(* IEC 61131-3 sources: daoli-st-library/DL_Algo (part 24) *)

(* ---- FB_DL_FoulingResistanceEstimator.st ---- *)
(*==============================================================================
 * 组件名称 (Component)  : FB_DL_FoulingResistanceEstimator
 * 所属子库 (Sublibrary) : DL_Algo
 * 当前版本 (Version)    : 1.0.0
 * 组件分类 (Category)   : 功能块（FUNCTION_BLOCK）· 换热器本体退化算法底座
 * 兼容性   (Platform)   : CODESYS 3.5 / TwinCAT 3 / 汇川 InoProShop / Schneider Machine Expert
 *                         仅依赖 Standard.library（R_TRIG / LN / ABS / MIN / MAX / LIMIT），零厂商方言
 * 接口依赖 (Depends)    : E_DL_Ne107Status —— 唯一属主为 DL_Device 子库的契约件
 *                         I_DL_DeviceHealth（R13 泳道 A1）。本文件只按成员名引用该枚举，
 *                         不重复定义枚举体（重复定义即同名异型，R33 家族超集风险）。
 * 功能描述 (Function)   : 由热侧/冷侧进出口温度与体积流量算出换热量 Q、对数平均温差
 *                         LMTD 与实测传热系数 K，再由 K 与清洁态基准 K_clean 反算污垢
 *                         热阻 Rf = 1/K − 1/K_clean；在趋势窗 tWindow 内用最小二乘做
 *                         Rf 对时间的线性拟合，输出增长斜率与清洗建议。
 *                         本件是「换热器污垢趋势」工艺件的算法底座：只做「算一个值 +
 *                         算一个趋势」，不判工艺合格、不控阀门、不做结垢成分分析。
 * 边界     (Boundary)   : ① 不做 PID、不做阀门/泵控制；② 不做结垢成分与化学分析；
 *                         ③ 数据不可信（温差过小 / 流量过低 / 两侧热负荷不平衡 /
 *                            输入非有限）时**拒绝更新**并保持上次有效值 —— 宁可不给
 *                            数，也不给脏数（R42 精神：判可用与取值同拍）；
 *                         ④ 不内置换热器几何模型与介质物性库，fCp/fRho 与 K_clean 全部
 *                            由调用方按设备台账注入。
 * 分层声明 (Layer)      : 算法层（DL_Algo）。上游为工艺台账件与 HMI 趋势，下游仅
 *                         Standard.library。零全局变量表引用、零外部变量声明、零物理 IO。
 * 段序     (Segments)   : 段1 实例无条件刷新 → 段2 复位通道（CASE 之前，R39）→
 *                         段3 参数闸门与输入防御 → 段4 数据质量四判据 → 段5 状态机 →
 *                         段6 有效更新与趋势累计 → 段7 结论仲裁 → 段8 码位单一优先级链 →
 *                         段9 出口钳位与保持语义重写。
 * 枚举映射表 (R31)      : eIdle(0)→标签 0｜eValid(10)→标签 10｜eTrend(20)→标签 20｜
 *                         eAdvice(30)→标签 30｜eFault(99)→标签 99。每个成员有且仅有一个
 *                         显式标签，ELSE 只接脏值（2212）。
 * 单拍标志清单 (R25)    : 本件唯一的沿输入是 bReset（复位），其消费点为段2 复位通道。
 *                         预清零点：段1 末（_bResetEdge := _fbTrigReset.Q 每次覆盖）；
 *                         置位点：段1 的 _fbTrigReset 实例调用；自清点：紧随实例调用之后
 *                         的 _bResetEdge 赋值行（下拍 R_TRIG.Q 转假即自然清）。
 * 保持位清单 (R27)      : bCleanAdvice（清洗建议，逐拍由 _bCleanLatched 重写）｜
 *                         fQ / fLmtd / fK / fRf（上次有效值，逐拍由 _fXxxHeld 重写并钳位）｜
 *                         fRfSlope（上次窗口斜率，逐拍重写）。复位沿清除锁存与保持值。
 * 定时器清单 (R40)      : 无 TON/TOF 实例。趋势窗以引脚 tSamplePeriod 累加计时，
 *                         窗边界显式重装基准（_fWinElapsedH := 0），不存在跨窗恒真输入；
 *                         时长到**或**样本数触顶（64）即结算并重开新窗，触顶提前结算是为了
 *                         避免「为了凑时长而丢掉分辨率」，也避免样本触顶后窗永远关不上。
 * 三元一致表 (R35)      : 流量比例守卫 0.05~0.9 / 封顶 0.9 / 判据 `<`（低于即不更新）｜
 *                         热平衡容差守卫 0.02~0.5 / 封顶 0.5 / 判据 `>`（超出即不更新）｜
 *                         最小温差守卫 0.5~20 K / 封顶 20 K / 判据 `<`（低于即不更新）。
 * 镜像量清单 (R38)      : 实时量 fFlowHot / fFlowCold 的唯一消费点是段4 的流量比例
 *                         判定（自学习参考流量 _fFlowHotMax / _fFlowColdMax 在同段更新）；
 *                         本件不设「锁存副本 + 实时镜像」双源，边界量全部取自本拍单次读取。
 * 开源溯源 (Origin)     : 原创实现（参考 OSCAT Building 的「温度/流量进 → 传热系数与
 *                         污垢热阻出」行为定义组织方式，T1-2；OSCAT 现行版为 EPL-2.0，
 *                         归档旧件仍受其原始许可约束 —— 本件只取行为定义与引脚组织，
 *                         未下载库文件、未复制任何源码行，公式取自公开传热学常识：
 *                         Q = m·cp·ΔT、逆/顺流 LMTD、Rf = 1/K − 1/K_clean）。
 *                         许可证结论：无代码复制，本文件为本库原创，随本库许可证发布。
 * 验收向量 (Acceptance) :
 *   V1 热侧 90/70 ℃、冷侧 20/40 ℃、逆流、两侧 10 m³/h：ΔT1 = 90−40 = 50 K、
 *      ΔT2 = 70−20 = 50 K，两温差相等时 LMTD 退化为算术平均 50.0 K；fQ ≈ 232.2 kW
 *      （10 m³/h × 1000 kg/m³ × 4.18 kJ/(kg·K) × 20 K / 3600）。规格记 49.7 K 与
 *      232 kW 为取整口径，本件按上式复算（见偏离留档②）。
 *   V2 fK = 1000、fKClean = 2000 → fRf = 1/1000 − 1/2000 = 5.0E-4 ≥ 3.0E-4 →
 *      bCleanAdvice = TRUE（保持态逐拍重写）。
 *   V3（V-A 除零）fArea = 0 → 16#0002_2210，fK 保持上次值并夹进 ≥ 0（R43）。
 *   V4（V-C 跨拍复验）进入 eTrend 后当拍流量骤降 → 段4 本拍复验流量门限失败 →
 *      本拍不更新、不累计斜率样本（绝不用上一相结论直接算斜率，R42）。
 *   V5（V-D 首拍）上电首拍 bValid = FALSE、fRf = 0.0，且首拍样本**不**写入趋势基准
 *      （R19：首扫只装基准，不参与斜率）。
 * 偏离留档 (Deviation)  :
 *   ① 「流量低于额定比例」的额定量：规格未给出额定流量引脚。本件以块内自学习的
 *      「投运以来观测到的最大流量」为参考（_fFlowHotMax / _fFlowColdMax），比例 =
 *      本拍流量 / 参考流量。理由：不新增引脚即可表达「相对自身额定」的语义；影响：
 *      上电初期参考流量偏低，门限自然宽松，随运行收敛（首拍样本不受门限影响）。
 *   ② V1 的 LMTD 数值：等温差时 LMTD 退化为算术平均（数值稳定性要求），与规格
 *      49.7 K 的取整口径相差 0.3 K，属口径差异而非算法差异，此处显式留档。
 *   ③ 输入非有限与「面积/清洁 K 非正」共用 16#0002_2210（规格故障表只给 3 个故障码，
 *      不新增码位；码位表以 §3.0 为准，编码者不得自行偏移）。
 * 修订历史 (Revision)   :
 *   2026-11-15  v1.0.0  首版入库（Round 13 · 泳道 C · DL_Algo 第 28 件）
 *============================================================================*)

(*-----------------------------------------------------------------------------
 * 枚举: E_DL_FoulingState（归属 FB_DL_FoulingResistanceEstimator，同文件发布）
 *----------------------------------------------------------------------------*)
TYPE E_DL_FoulingState :
(
    eIdle   := 0,    // 空闲：未使能或参数未就绪 / Idle, disabled or parameters not ready
    eValid  := 10,   // 有效：本拍已算出可信的 K 与 Rf / Valid, trustworthy K and Rf computed
    eTrend  := 20,   // 趋势：窗内样本数已达 3，斜率可算 / Trend, at least three window samples
    eAdvice := 30,   // 建议清洗：热阻或其斜率越阈（锁存）/ Cleaning advised, latched
    eFault  := 99    // 故障：参数非法或输入非有限 / Fault, illegal parameter or non-finite input
) UINT;
END_TYPE

FUNCTION_BLOCK FB_DL_FoulingResistanceEstimator
VAR_INPUT
    bEnable         : BOOL;                 // 使能（Enable），FALSE = 冻结更新并回空闲；复位通道不受其屏蔽 / Enable, FALSE freezes updates
    bReset          : BOOL;                 // 复位（Reset），上升沿清趋势窗、清洗锁存与保持值 / Rising edge clears trend window and latches
    fTinHot         : REAL;                 // 热侧进口温度（Hot inlet temperature）[℃]，域 −50~300 / Hot side inlet temperature [degC]
    fToutHot        : REAL;                 // 热侧出口温度（Hot outlet temperature）[℃]，域 −50~300 / Hot side outlet temperature [degC]
    fTinCold        : REAL;                 // 冷侧进口温度（Cold inlet temperature）[℃]，域 −50~300 / Cold side inlet temperature [degC]
    fToutCold       : REAL;                 // 冷侧出口温度（Cold outlet temperature）[℃]，域 −50~300 / Cold side outlet temperature [degC]
    fFlowHot        : REAL;                 // 热侧体积流量（Hot volumetric flow）[m³/h]，域 0~10000 / Hot volumetric flow [m3/h]
    fFlowCold       : REAL;                 // 冷侧体积流量（Cold volumetric flow）[m³/h]，域 0~10000 / Cold volumetric flow [m3/h]
    fCpHot          : REAL := 4.18;         // 热侧比热（Hot specific heat）[kJ/(kg·K)]，域 0.5~10，默认 4.18 / Hot specific heat [kJ/(kg K)]
    fCpCold         : REAL := 4.18;         // 冷侧比热（Cold specific heat）[kJ/(kg·K)]，域 0.5~10，默认 4.18 / Cold specific heat [kJ/(kg K)]
    fRhoHot         : REAL := 1000.0;       // 热侧密度（Hot density）[kg/m³]，域 1~2000，默认 1000.0 / Hot density [kg/m3]
    fRhoCold        : REAL := 1000.0;       // 冷侧密度（Cold density）[kg/m³]，域 1~2000，默认 1000.0 / Cold density [kg/m3]
    fArea           : REAL;                 // 换热面积（Heat transfer area）[m²]，域 >0，除零保护对象 / Heat transfer area [m2], must be positive
    fKClean         : REAL;                 // 清洁态传热系数基准（Clean-condition K）[W/(m²·K)]，域 >0 / Clean-condition K [W/(m2 K)], must be positive
    bCounterFlow    : BOOL := TRUE;         // 流型（Flow arrangement），TRUE = 逆流，FALSE = 顺流，默认 TRUE / TRUE counter-flow, FALSE parallel-flow
    fDtmMin         : REAL := 2.0;          // 最小可用温差（Minimum usable temperature difference）[K]，域 0.5~20，默认 2.0 / Minimum usable LMTD [K]
    fHeatBalTol     : REAL := 0.10;         // 两侧热负荷允许偏差比（Heat balance tolerance）[-]，域 0.02~0.5，默认 0.10 / Heat balance tolerance [-]
    fFlowMinRatio   : REAL := 0.20;         // 流量下限比例（Minimum flow ratio）[-]，域 0.05~0.9，默认 0.20 / Minimum flow ratio [-]
    tWindow         : TIME := T#1H;         // 趋势窗长（Trend window），域 5 min~24 h，默认 1 h / Trend window, default 1 h
    tSamplePeriod   : TIME := T#10S;        // 调用周期（Call period）[ms]，必须与实际任务周期一致，默认 10 s / Call period, must match the task
    fRfAlarm        : REAL := 3.0E-4;       // 污垢热阻报警阈（Fouling resistance alarm）[m²·K/W]，域 1E-5~5E-3 / Fouling resistance alarm [m2 K/W]
    fSlopeAlarm     : REAL := 2.0E-5;       // 污垢增长速率阈（Fouling slope alarm）[m²·K/(W·h)]，域 1E-7~1E-3 / Fouling slope alarm [m2 K/(W h)]
END_VAR

VAR_OUTPUT
    fQ              : REAL;                 // 热负荷两侧平均（Heat duty, mean of both sides）[kW]，保持语义 / Mean heat duty of both sides [kW], held
    fLmtd           : REAL;                 // 对数平均温差（Log mean temperature difference）[K]，保持语义 / LMTD [K], held
    fK              : REAL;                 // 实测传热系数（Measured overall K）[W/(m²·K)]，保持语义且夹进 ≥0 / Measured K [W/(m2 K)], held and clamped non-negative
    fRf             : REAL;                 // 污垢热阻（Fouling resistance）[m²·K/W]，= 1/K − 1/K_clean，保持语义 / Fouling resistance [m2 K/W], held
    fRfSlope        : REAL;                 // 窗内趋势斜率（Trend slope in window）[m²·K/(W·h)]，保持语义 / Trend slope [m2 K/(W h)], held
    bValid          : BOOL;                 // 本拍输出有效（Output valid this scan），数据质量不足时为 FALSE / TRUE when this scan produced a trustworthy value
    bCleanAdvice    : BOOL;                 // 建议清洗（Cleaning advised），保持语义（R27），复位沿清除 / Cleaning advised, held until reset
    eHealth         : E_DL_Ne107Status;     // 健康态（NE107 health），引用属主 A1 的枚举 / NE107 health state, owned by A1
    uDiagCode       : UDINT;                // 诊断码（Diagnostic code），本拍单一优先级链输出 / Diagnostic code, single priority chain
    uErrorId        : UDINT;                // 故障码（Error code），仅故障级码，0 = 无故障 / Fault-level code, 0 = no fault
    bError          : BOOL;                 // 故障标志（Error），仅故障级码置位，信息级不置位 / TRUE only for fault-level codes
    nUpdateCount    : UDINT;                // 有效更新次数（Valid update counter）[次]，每次有效更新 +1 / Valid update counter [count]
END_VAR

VAR
    _eState         : E_DL_FoulingState := E_DL_FoulingState.eIdle; // 内部状态（Internal state）/ Internal state machine value
    _bInit          : BOOL;                 // 首扫标志（First-scan flag），初值 FALSE，唯一首扫判据为 NOT _bInit（R19）/ First-scan flag, FALSE by default
    _bSkipSample    : BOOL;                 // 本拍不参与斜率（Skip trend sample this scan），首扫与不可信拍置位 / Skip this scan as a trend sample
    _bParamOk       : BOOL;                 // 参数闸门通过（Parameter gate passed）/ Parameter gate result
    _bDataOk        : BOOL;                 // 数据质量通过（Data quality passed）/ Data quality result
    _bValidNow      : BOOL;                 // 本拍有效（Valid this scan）/ Valid this scan
    _bFaultCond     : BOOL;                 // 故障条件（Fault condition latch-free flag）/ Fault condition flag
    _uFaultCode     : UDINT;                // 本拍故障级码（Fault-level code this scan）/ Fault-level code of this scan
    _uFaultLatched  : UDINT;                // 故障码锁存（Latched fault code），仅复位沿清除 / Latched fault code, reset only
    _uInfoCode      : UDINT;                // 本拍信息级码（Info-level code this scan），每拍重算 / Info-level code, recomputed every scan
    _bArrPrev       : BOOL;                 // 上拍流型（Previous flow arrangement）/ Flow arrangement of the previous scan
    _bArrKnown      : BOOL;                 // 流型已记录（Arrangement recorded）/ Arrangement recorded flag
    _fAreaEff       : REAL;                 // 生效换热面积（Effective area）[m²]，闸门后值 / Effective area [m2] after the gate
    _fKCleanEff     : REAL;                 // 生效清洁 K（Effective clean K）[W/(m²·K)] / Effective clean K [W/(m2 K)]
    _fDtmMinEff     : REAL;                 // 生效最小温差（Effective minimum LMTD）[K]，钳位 0.5~20 / Effective minimum LMTD [K], clamped
    _fBalTolEff     : REAL;                 // 生效热平衡容差（Effective heat balance tolerance）[-]，钳位 0.02~0.5 / Effective heat balance tolerance, clamped
    _fFlowRatioEff  : REAL;                 // 生效流量比例（Effective minimum flow ratio）[-]，钳位 0.05~0.9 / Effective minimum flow ratio, clamped
    _fFlowHotMax    : REAL;                 // 热侧参考流量（Hot reference flow）[m³/h]，自学习峰值 / Self-learned hot reference flow [m3/h]
    _fFlowColdMax   : REAL;                 // 冷侧参考流量（Cold reference flow）[m³/h]，自学习峰值 / Self-learned cold reference flow [m3/h]
    _fQHot          : REAL;                 // 热侧放热量（Heat duty, hot side）[kW]，有符号 / Hot-side duty [kW], signed
    _fQCold         : REAL;                 // 冷侧吸热量（Heat duty, cold side）[kW]，有符号 / Cold-side duty [kW], signed
    _fQMean         : REAL;                 // 两侧平均热负荷（Mean duty）[kW] / Mean duty of both sides [kW]
    _fDt1           : REAL;                 // 端差一（Terminal difference one）[K]，按流型取 / Terminal temperature difference one [K]
    _fDt2           : REAL;                 // 端差二（Terminal difference two）[K]，按流型取 / Terminal temperature difference two [K]
    _fLmtdCalc      : REAL;                 // 本拍 LMTD 计算值（Computed LMTD）[K] / Computed LMTD [K]
    _fLmtdAbs       : REAL;                 // 端差差值的绝对值（Absolute terminal difference gap）[K]，退化判据 / Absolute gap between terminal differences [K]
    _fLmtdDen       : REAL;                 // 对数比值（Logarithmic ratio）[-]，除零保护对象 / Logarithmic ratio, divide-guard object
    _fBalDev        : REAL;                 // 热平衡偏差比（Heat balance deviation）[-] / Heat balance deviation ratio [-]
    _fBalRef        : REAL;                 // 热平衡参考量（Heat balance reference）[kW]/ Reference magnitude for the balance test [kW]
    _fKCalc         : REAL;                 // 本拍 K 计算值（Computed K）[W/(m²·K)] / Computed K [W/(m2 K)]
    _fRfCalc        : REAL;                 // 本拍 Rf 计算值（Computed Rf）[m²·K/W] / Computed Rf [m2 K/W]
    _fQHeld         : REAL;                 // 保持的热负荷（Held heat duty）[kW] / Held heat duty [kW]
    _fLmtdHeld      : REAL;                 // 保持的 LMTD（Held LMTD）[K] / Held LMTD [K]
    _fKHeld         : REAL;                 // 保持的 K（Held K）[W/(m²·K)] / Held K [W/(m2 K)]
    _fRfHeld        : REAL;                 // 保持的 Rf（Held Rf）[m²·K/W] / Held Rf [m2 K/W]
    _fSlopeHeld     : REAL;                 // 保持的斜率（Held slope）[m²·K/(W·h)] / Held slope [m2 K/(W h)]
    _bCleanLatched  : BOOL;                 // 清洗建议锁存（Cleaning advice latch），仅复位沿清除 / Cleaning advice latch, reset only
    _nWinN          : INT;                  // 窗内样本数（Window sample count）[个]，上限 64 / Window sample count, capped at 64
    _fWinElapsedH   : REAL;                 // 窗内已历时（Elapsed hours in window）[h] / Elapsed hours in the current window [h]
    _fWinX          : REAL;                 // 最小二乘 Σt（Sum of time stamps）[h] / Least-squares sum of time stamps [h]
    _fWinY          : REAL;                 // 最小二乘 ΣRf（Sum of Rf samples）[m²·K/W] / Least-squares sum of Rf samples [m2 K/W]
    _fWinXY         : REAL;                 // 最小二乘 Σt·Rf（Sum of products）[h·m²·K/W] / Least-squares sum of products
    _fWinXX         : REAL;                 // 最小二乘 Σt²（Sum of squared times）[h²] / Least-squares sum of squared times [h2]
    _fWinDen        : REAL;                 // 最小二乘分母（Normal-equation denominator）[-]，除零保护对象 / Denominator of the normal equations
    _fWinNum        : REAL;                 // 最小二乘分子（Normal-equation numerator）[-] / Numerator of the normal equations
    _fDtHours       : REAL;                 // 本拍步长（Step in hours）[h]，由 tSamplePeriod 折算 / Step in hours, derived from the call period
    _fWinHoursEff   : REAL;                 // 生效窗长（Effective window length）[h]，由 tWindow 折算 / Effective window length [h]
    _fbTrigReset    : R_TRIG;               // 复位沿（Reset edge detector），主体最前部无条件刷新 / Reset edge detector, refreshed unconditionally
    _bResetEdge     : BOOL;                 // 复位沿单拍标志（Reset one-shot flag），紧随实例自清 / Reset one-shot flag, cleared right after the call
END_VAR

VAR CONSTANT
    DL_FRE_REAL_MAX   : REAL := 3.4E38;      // 单精度有限值判据幅值（Finite magnitude bound）/ Finite bound for REAL inputs
    DL_FRE_EPS        : REAL := 1.0E-6;      // 浮点防零容差（Divide-guard epsilon）/ Float divide-guard epsilon
    DL_FRE_K_MAX      : REAL := 1.0E9;       // K 出口上限（K output ceiling）[W/(m²·K)] / Upper clamp of K [W/(m2 K)]
    DL_FRE_RF_MAX     : REAL := 1.0;         // Rf 出口上限（Rf output ceiling）[m²·K/W] / Upper clamp of Rf [m2 K/W]
    DL_FRE_SLOPE_MAX  : REAL := 1.0;         // 斜率出口上限（Slope output ceiling）[m²·K/(W·h)] / Upper clamp of slope
    DL_FRE_SLOPE_MIN  : REAL := -1.0;        // 斜率出口下限（Slope output floor）[m²·K/(W·h)] / Lower clamp of slope
    DL_FRE_WIN_MAX    : INT  := 64;          // 窗内样本上限（Window sample ceiling）[个] / Window sample ceiling
    DL_FRE_MS_PER_H   : REAL := 3600000.0;   // 毫秒→小时换算（Milliseconds-to-hours scale）[-] / Milliseconds-to-hours scale
    DL_FRE_KW_SCALE   : REAL := 3600.0;      // m³/h·kg/m³·kJ/(kg·K)·K → kW 的换算（Duty unit scale）[-] / Duty unit scale
    DL_FRE_W_SCALE    : REAL := 1000.0;      // kW → W 换算（Kilowatt-to-watt scale）[-] / Kilowatt-to-watt scale
    DL_FRE_DTM_MIN    : REAL := 0.5;         // 最小温差域下限（Minimum LMTD lower clamp）[K] / Minimum LMTD lower clamp [K]
    DL_FRE_DTM_MAX    : REAL := 20.0;        // 最小温差域上限（Minimum LMTD upper clamp）[K] / Minimum LMTD upper clamp [K]
    DL_FRE_TOL_MIN    : REAL := 0.02;        // 热平衡容差域下限（Balance tolerance lower clamp）[-] / Balance tolerance lower clamp
    DL_FRE_TOL_MAX    : REAL := 0.5;         // 热平衡容差域上限（Balance tolerance upper clamp）[-] / Balance tolerance upper clamp
    DL_FRE_RATIO_MIN  : REAL := 0.05;        // 流量比例域下限（Flow ratio lower clamp）[-] / Flow ratio lower clamp
    DL_FRE_RATIO_MAX  : REAL := 0.9;         // 流量比例域上限（Flow ratio upper clamp）[-] / Flow ratio upper clamp
    DL_FRE_RF_FLOOR   : REAL := 0.0;         // Rf 出口下限（Rf output floor）[m²·K/W]，K>K_clean 时按 0 / Rf floor, zero when K exceeds clean K
    DL_FRE_WIN_MIN_N  : INT  := 3;           // 斜率所需最少样本（Minimum samples for a slope）[个] / Minimum samples for the slope
    DL_FRE_ERR_PARAM  : UDINT := 16#0002_2210; // 0002_2210 面积/清洁 K 非正或输入非有限【故障级】/ Illegal area, clean K or non-finite input
    DL_FRE_ERR_LMTD   : UDINT := 16#0002_2211; // 0002_2211 LMTD ≤ 0（温度交叉或流型用错）【故障级】/ Non-positive LMTD
    DL_FRE_ERR_STATE  : UDINT := 16#0002_2212; // 0002_2212 非法状态兜底【故障级】/ Illegal state fallback
    DL_FRE_INFO_LMTD  : UDINT := 16#0002_2201; // 0002_2201 LMTD 低于最小可用温差【信息级】/ LMTD below the usable limit
    DL_FRE_INFO_FLOW  : UDINT := 16#0002_2202; // 0002_2202 流量低于下限比例【信息级】/ Flow below the minimum ratio
    DL_FRE_INFO_BAL   : UDINT := 16#0002_2203; // 0002_2203 两侧热负荷偏差超容差【信息级】/ Heat balance exceeded
    DL_FRE_INFO_ARR   : UDINT := 16#0002_2204; // 0002_2204 逆/顺流口径切换，趋势基准已重置【信息级】/ Arrangement changed, trend reset
END_VAR

// ============================================================================
// 段 1｜实例无条件周期刷新（R7/0.5：严禁置于 IF / CASE 分支内）
//      Unconditional per-cycle refresh of every instance (R7/0.5)
// ============================================================================
_fbTrigReset(CLK := bReset);            // 复位沿实例调用（Reset edge instance call）
_bResetEdge := _fbTrigReset.Q;          // 单拍标志紧随实例赋值，下拍自然清（R24/R25 自清点）

// 本拍故障/信息码与结论预置（每拍重算，杜绝跨拍残留）
// Per-scan preset of codes and conclusions, no cross-scan residue
_uFaultCode  := _uFaultLatched;         // 故障码以上拍锁存续用（Carry the latched fault code）
_uInfoCode   := 16#0000_0000;           // 信息级码预清零（Info code preset to zero）
_bFaultCond  := FALSE;                  // 故障条件预清零（Fault condition preset FALSE）
_bParamOk    := FALSE;                  // 参数闸门预置未通过（Parameter gate preset closed）
_bDataOk     := FALSE;                  // 数据质量预置未通过（Data quality preset failed）
_bValidNow   := FALSE;                  // 本拍有效预置假（Valid preset FALSE）
_bSkipSample := FALSE;                  // 采样跳过预置假（Sample skip preset FALSE）

// 调用周期折算为小时，非法周期按复位通道外的钳位处理（不做除零）
// Convert the call period into hours, illegal periods are clamped instead of divided by zero
IF tSamplePeriod >= T#1MS THEN
    _fDtHours := TIME_TO_REAL(tSamplePeriod) / DL_FRE_MS_PER_H;   // 毫秒 → 小时（Milliseconds to hours）
ELSE
    _fDtHours := 0.0;                   // 周期非法时不推进窗口（Illegal period does not advance the window）
    _bFaultCond := TRUE;                // 周期非法按参数故障处理（Illegal period treated as a parameter fault）
    _uFaultCode := DL_FRE_ERR_PARAM;    // 0002_2210 周期非法并入参数故障【故障级】/ Illegal period folded into the parameter fault
END_IF

// ============================================================================
// 段 2｜复位通道（R39：置于 CASE 之前，且不被掉使能分支屏蔽）
//      Reset path, placed before CASE and never masked by the disable branch
// ============================================================================
IF _bResetEdge THEN
    _bCleanLatched := FALSE;            // 清洗建议锁存清除（Cleaning advice latch cleared）
    _nWinN         := 0;                // 窗内样本数清零（Window sample count cleared）
    _fWinElapsedH  := 0.0;              // 窗内历时清零（Window elapsed cleared）
    _fWinX         := 0.0;              // Σt 清零（Sum of time cleared）
    _fWinY         := 0.0;              // ΣRf 清零（Sum of Rf cleared）
    _fWinXY        := 0.0;              // Σt·Rf 清零（Sum of products cleared）
    _fWinXX        := 0.0;              // Σt² 清零（Sum of squares cleared）
    _fSlopeHeld    := 0.0;              // 斜率保持值清零（Held slope cleared）
    _fRfHeld       := 0.0;              // Rf 保持值清零（Held Rf cleared）
    _fKHeld        := 0.0;              // K 保持值清零（Held K cleared）
    _fQHeld        := 0.0;              // 热负荷保持值清零（Held duty cleared）
    _fLmtdHeld     := 0.0;              // LMTD 保持值清零（Held LMTD cleared）
    _uFaultLatched := 16#0000_0000;     // 故障码锁存清除（Latched fault code cleared）
    _uFaultCode    := 16#0000_0000;     // 本拍故障码随复位清空，防止段8 重新锁存旧码（Clear this scan code）
    IF _eState = E_DL_FoulingState.eFault THEN
        _eState := E_DL_FoulingState.eIdle;  // 故障态回空闲（Fault state back to idle）
        _uFaultCode := 16#0000_0000;    // 故障码随复位清除（Fault code cleared with the reset）
        _bFaultCond := FALSE;           // 故障条件随复位清除（Fault condition cleared）
    END_IF
END_IF

// ============================================================================
// 段 3｜参数闸门与输入防御（先判可用，再算值；R42 同源纪律）
//      Parameter gate and input defense: availability first, arithmetic second
// ============================================================================
IF (NOT (fArea     >= (-DL_FRE_REAL_MAX) AND fArea     <= DL_FRE_REAL_MAX))
OR (NOT (fKClean   >= (-DL_FRE_REAL_MAX) AND fKClean   <= DL_FRE_REAL_MAX))
OR (NOT (fTinHot   >= (-DL_FRE_REAL_MAX) AND fTinHot   <= DL_FRE_REAL_MAX))
OR (NOT (fToutHot  >= (-DL_FRE_REAL_MAX) AND fToutHot  <= DL_FRE_REAL_MAX))
OR (NOT (fTinCold  >= (-DL_FRE_REAL_MAX) AND fTinCold  <= DL_FRE_REAL_MAX))
OR (NOT (fToutCold >= (-DL_FRE_REAL_MAX) AND fToutCold <= DL_FRE_REAL_MAX))
OR (NOT (fFlowHot  >= (-DL_FRE_REAL_MAX) AND fFlowHot  <= DL_FRE_REAL_MAX))
OR (NOT (fFlowCold >= (-DL_FRE_REAL_MAX) AND fFlowCold <= DL_FRE_REAL_MAX))
OR (NOT (fCpHot    >= (-DL_FRE_REAL_MAX) AND fCpHot    <= DL_FRE_REAL_MAX))
OR (NOT (fCpCold   >= (-DL_FRE_REAL_MAX) AND fCpCold   <= DL_FRE_REAL_MAX))
OR (NOT (fRhoHot   >= (-DL_FRE_REAL_MAX) AND fRhoHot   <= DL_FRE_REAL_MAX))
OR (NOT (fRhoCold  >= (-DL_FRE_REAL_MAX) AND fRhoCold  <= DL_FRE_REAL_MAX))
OR (NOT (fRfAlarm  >= (-DL_FRE_REAL_MAX) AND fRfAlarm  <= DL_FRE_REAL_MAX))
OR (NOT (fSlopeAlarm >= (-DL_FRE_REAL_MAX) AND fSlopeAlarm <= DL_FRE_REAL_MAX)) THEN
    _bFaultCond := TRUE;                // 任一输入非有限即故障（Any non-finite input is a fault）
    _uFaultCode := DL_FRE_ERR_PARAM;    // 0002_2210 输入非有限【故障级】/ Non-finite input, fault level
ELSIF fArea <= 0.0 THEN
    _bFaultCond := TRUE;                // 面积非正：K 的分母不可用（Non-positive area breaks the K denominator）
    _uFaultCode := DL_FRE_ERR_PARAM;    // 0002_2210 面积非正【故障级】/ Illegal area, fault level
ELSIF fKClean <= 0.0 THEN
    _bFaultCond := TRUE;                // 清洁 K 非正：Rf 的基准不可用（Non-positive clean K breaks the Rf basis）
    _uFaultCode := DL_FRE_ERR_PARAM;    // 0002_2210 清洁 K 非正【故障级】/ Illegal clean K, fault level
ELSE
    _bParamOk := TRUE;                  // 参数闸门通过（Parameter gate passed）
END_IF

// 生效参数的域钳位（R35：守卫、封顶值、判据运算符三者同向）
// Clamp effective parameters, keeping guard, ceiling and comparison operator in step (R35)
_fDtmMinEff    := LIMIT(DL_FRE_DTM_MIN, fDtmMin, DL_FRE_DTM_MAX);       // 最小温差钳位 0.5~20 K（Minimum LMTD clamped）
_fBalTolEff    := LIMIT(DL_FRE_TOL_MIN, fHeatBalTol, DL_FRE_TOL_MAX);   // 热平衡容差钳位 0.02~0.5（Balance tolerance clamped）
_fFlowRatioEff := LIMIT(DL_FRE_RATIO_MIN, fFlowMinRatio, DL_FRE_RATIO_MAX); // 流量比例钳位 0.05~0.9（Flow ratio clamped）
_fWinHoursEff  := TIME_TO_REAL(tWindow) / DL_FRE_MS_PER_H;   // 窗长折算为小时（Window length in hours）
_fAreaEff      := fArea;                // 面积已过正数防御（Area already defended positive inside the gate）
_fKCleanEff     := fKClean;             // 清洁 K 已过正数防御（Clean K already defended positive inside the gate）

// 参考流量自学习（偏离留档①）：上电初期参考值随运行收敛，仅用于相对流量判定
// Self-learned reference flow (deviation 1): converges during commissioning, used for the relative flow test
IF fFlowHot >= 0.0 THEN
    _fFlowHotMax  := MAX(_fFlowHotMax, fFlowHot);   // 热侧参考取历史峰值（Hot reference takes the historic peak）
ELSE
    _fFlowHotMax  := _fFlowHotMax;                  // 负流量不参与自学习（Negative flow is not learned）
END_IF
IF fFlowCold >= 0.0 THEN
    _fFlowColdMax := MAX(_fFlowColdMax, fFlowCold); // 冷侧参考取历史峰值（Cold reference takes the historic peak）
ELSE
    _fFlowColdMax := _fFlowColdMax;                 // 负流量不参与自学习（Negative flow is not learned）
END_IF

// ============================================================================
// 段 4｜数据质量四判据（本拍复验；判「可用」与取「值」同拍完成，R42）
//      Four data-quality criteria, all re-evaluated on this very scan (R42)
// ============================================================================
IF _bParamOk AND bEnable AND (NOT _bFaultCond) THEN

    // 4.1 计算两侧热负荷（有符号，kW）：Q = V̇ · ρ · cp · ΔT / 3600
    //     Duty on both sides, signed, in kW
    _fQHot  := fFlowHot  * fRhoHot  * fCpHot  * (fTinHot  - fToutHot)  / DL_FRE_KW_SCALE;
    _fQCold := fFlowCold * fRhoCold * fCpCold * (fToutCold - fTinCold) / DL_FRE_KW_SCALE;
    _fQMean := (ABS(_fQHot) + ABS(_fQCold)) / 2.0;   // 两侧平均热负荷（Mean duty of both sides）

    // 4.2 端差按流型取：逆流对热进-冷出；顺流对热进-冷进
    //     Terminal differences by flow arrangement
    IF bCounterFlow THEN
        _fDt1 := fTinHot - fToutCold;   // 逆流端差一（Counter-flow terminal difference one）
        _fDt2 := fToutHot - fTinCold;   // 逆流端差二（Counter-flow terminal difference two）
    ELSE
        _fDt1 := fTinHot - fTinCold;    // 顺流端差一（Parallel-flow terminal difference one）
        _fDt2 := fToutHot - fToutCold;  // 顺流端差二（Parallel-flow terminal difference two）
    END_IF

    // 4.3 LMTD：端差相等时退化为算术平均，避免 ln(1)=0 造成除零
    //     LMTD degenerates to the arithmetic mean when both terminal differences are equal
    _fLmtdAbs := ABS(_fDt1 - _fDt2);    // 端差差值绝对值（Absolute gap of the terminal differences）
    IF _fLmtdAbs < DL_FRE_EPS THEN
        _fLmtdCalc := (_fDt1 + _fDt2) / 2.0;    // 等温差退化（Equal-difference degeneration）
    ELSIF (_fDt1 <= 0.0) OR (_fDt2 <= 0.0) THEN
        _fLmtdCalc := 0.0;              // 温度交叉：本拍不可算（Temperature cross, not computable）
    ELSE
        _fLmtdDen  := _fDt1 / _fDt2;    // 对数比值（Logarithmic ratio），两端差均为正才有意义
        _fLmtdCalc := (_fDt1 - _fDt2) / LN(_fLmtdDen);   // 标准 LMTD 定义（Standard LMTD definition）
    END_IF

    // 4.4 流型切换：趋势基准必须重置，否则跨流型样本混算斜率
    //     Arrangement change forces a trend reset, mixing arrangements would corrupt the slope
    IF _bArrKnown AND (bCounterFlow <> _bArrPrev) THEN
        _nWinN        := 0;             // 窗内样本清零（Window samples cleared）
        _fWinElapsedH := 0.0;           // 窗内历时清零（Window elapsed cleared）
        _fWinX        := 0.0;           // Σt 清零（Sum of time cleared）
        _fWinY        := 0.0;           // ΣRf 清零（Sum of Rf cleared）
        _fWinXY       := 0.0;           // Σt·Rf 清零（Sum of products cleared）
        _fWinXX       := 0.0;           // Σt² 清零（Sum of squares cleared）
        _uInfoCode    := DL_FRE_INFO_ARR;   // 0002_2204 流型切换趋势重置【信息级】/ Arrangement changed, info level
    END_IF
    _bArrPrev  := bCounterFlow;         // 记录本拍流型（Record this scan arrangement）
    _bArrKnown := TRUE;                 // 流型已记录（Arrangement recorded）

    // 4.5 四判据依次裁决：LMTD 非法 > 温差不足 > 流量不足 > 热平衡超差
    //     Four criteria in a single priority chain
    IF _fLmtdCalc <= 0.0 THEN
        _bFaultCond := TRUE;            // LMTD 非正属故障级（Non-positive LMTD is a fault）
        _uFaultCode := DL_FRE_ERR_LMTD; // 0002_2211 LMTD ≤ 0【故障级】/ Non-positive LMTD, fault level
    ELSIF _fLmtdCalc < _fDtmMinEff THEN
        _uInfoCode := DL_FRE_INFO_LMTD; // 0002_2201 温差太小不可信【信息级】/ LMTD below usable limit
    ELSIF (_fFlowHotMax > DL_FRE_EPS) AND ((fFlowHot / _fFlowHotMax) < _fFlowRatioEff) THEN
        _uInfoCode := DL_FRE_INFO_FLOW; // 0002_2202 热侧流量过低【信息级】/ Hot flow below the ratio
    ELSIF (_fFlowColdMax > DL_FRE_EPS) AND ((fFlowCold / _fFlowColdMax) < _fFlowRatioEff) THEN
        _uInfoCode := DL_FRE_INFO_FLOW; // 0002_2202 冷侧流量过低【信息级】/ Cold flow below the ratio
    ELSE
        _fBalRef := MAX(ABS(_fQHot), ABS(_fQCold));  // 热平衡参考量（Balance reference magnitude）
        IF _fBalRef > DL_FRE_EPS THEN
            _fBalDev := ABS(_fQHot - _fQCold) / _fBalRef;   // 偏差比（Deviation ratio）
        ELSE
            _fBalDev := 1.0;            // 两侧均为零：按最坏偏差处理（Both sides zero: worst case）
        END_IF
        IF _fBalDev > _fBalTolEff THEN
            _uInfoCode := DL_FRE_INFO_BAL;  // 0002_2203 热平衡超差【信息级】/ Heat balance exceeded
        ELSE
            _bDataOk := TRUE;           // 数据质量通过（Data quality passed）
        END_IF
    END_IF
END_IF

// ============================================================================
// 段 5｜状态机（ENUM + CASE，含 ELSE 非法状态兜底）
//      State machine with an explicit ELSE fallback
// ============================================================================
IF _bFaultCond THEN
    _eState := E_DL_FoulingState.eFault;    // 故障条件优先于状态机（Fault condition outranks the machine）
END_IF

// 掉使能冻结分支：显式排除故障态，复位通道仍可从故障态退出（R39 合法写法①）
// Disable branch explicitly excludes the fault state, the reset path still works (R39 form 1)
IF (NOT bEnable) AND (_eState <> E_DL_FoulingState.eFault) THEN
    _eState := E_DL_FoulingState.eIdle;     // 冻结回空闲（Freeze back to idle）
    _bDataOk := FALSE;                      // 掉使能时数据质量结论作废（Quality result voided while disabled）
END_IF

CASE _eState OF

    E_DL_FoulingState.eIdle: // 空闲：等使能与参数闸门
        IF bEnable AND _bParamOk AND (NOT _bFaultCond) THEN
            _eState := E_DL_FoulingState.eValid;    // 进有效态（Enter valid state）
        END_IF

    E_DL_FoulingState.eValid: // 有效：等待窗内样本积累
        IF _bDataOk AND (_nWinN >= DL_FRE_WIN_MIN_N) THEN
            _eState := E_DL_FoulingState.eTrend;    // 样本足够进趋势态（Enough samples, enter trend）
        END_IF

    E_DL_FoulingState.eTrend: // 趋势：持续累计，越阈转建议
        IF _bCleanLatched THEN
            _eState := E_DL_FoulingState.eAdvice;   // 越阈转建议清洗（Threshold crossed, advise cleaning）
        END_IF

    E_DL_FoulingState.eAdvice: // 建议清洗：锁存至复位，本分支只做出口重写（R27）
        // 结论与出口在本分支外逐拍重写，此处仅保留空标签与原因注释（R31）
        // Outputs are rewritten outside this branch every scan, so the label stays empty (R31)

    E_DL_FoulingState.eFault: // 故障：等复位沿
        // 复位通道位于 CASE 之前，本分支无需动作，保留标签与原因注释（R31/R39）
        // The reset path sits before CASE, so this branch only keeps the label (R31/R39)

    ELSE // 兜底：非法状态
        _uFaultCode := DL_FRE_ERR_STATE;        // 0002_2212 非法状态兜底【故障级】/ Illegal state fallback
        _bFaultCond := TRUE;                    // 置故障条件（Raise the fault condition）
        _eState     := E_DL_FoulingState.eFault;    // 强制回故障态（Force the fault state）
END_CASE

// ============================================================================
// 段 6｜有效更新与趋势累计（首扫只装基准，不参与斜率，R19）
//      Valid update and trend accumulation, the first scan only loads the basis (R19)
// ============================================================================
IF _bDataOk AND (_eState <> E_DL_FoulingState.eFault) THEN
    _fKCalc := (_fQMean * DL_FRE_W_SCALE) / (_fAreaEff * _fLmtdCalc);   // K = Q / (A · LMTD)
    _fRfCalc := 0.0;                    // Rf 预置 0（Rf preset to zero）
    IF _fKCalc > DL_FRE_EPS THEN
        _fRfCalc := (1.0 / _fKCalc) - (1.0 / _fKCleanEff);  // Rf = 1/K − 1/K_clean
    ELSE
        _fRfCalc := 0.0;                // K 过小按不可算处理（K too small, treated as not computable）
    END_IF
    IF _fRfCalc < DL_FRE_RF_FLOOR THEN
        _fRfCalc := DL_FRE_RF_FLOOR;    // 负污垢（比清洁态更好）按 0（Negative fouling floored to zero）
    END_IF

    // 首扫只装基准：本拍只把有效值写进保持量，不压入趋势样本（R19）
    // First scan loads the basis only: hold the value but never push a trend sample (R19)
    IF NOT _bInit THEN
        _bInit       := TRUE;           // 首扫完成（First scan done）
        _bSkipSample := TRUE;           // 本拍不参与斜率（Do not take a trend sample this scan）
    END_IF

    _fQHeld    := _fQMean;              // 热负荷保持（Duty held）
    _fLmtdHeld := _fLmtdCalc;           // LMTD 保持（LMTD held）
    _fKHeld    := _fKCalc;              // K 保持（K held）
    _fRfHeld   := _fRfCalc;             // Rf 保持（Rf held）
    nUpdateCount := nUpdateCount + UDINT#1; // 有效更新计数（Valid update counted）
    _bValidNow := TRUE;                 // 本拍有效（Valid this scan）

    // 趋势累计：窗内最小二乘（Σt、ΣRf、Σt·Rf、Σt²）
    // Trend accumulation with the normal-equation sums
    //   计时必须**无条件**推进：若只在压样本时才推进，样本数触顶后窗内历时停止增长，
    //   窗永远关不上，斜率也就永远算不出来（这是本件最容易写死的一处）。
    //   Elapsed time advances unconditionally, otherwise a capped sample count freezes the window.
    _fWinElapsedH := _fWinElapsedH + _fDtHours;         // 窗内历时推进（Window elapsed advances）
    IF (NOT _bSkipSample) AND (_nWinN < DL_FRE_WIN_MAX) THEN
        _fWinX        := _fWinX + _fWinElapsedH;        // Σt 累加（Sum of time accumulates）
        _fWinY        := _fWinY + _fRfCalc;             // ΣRf 累加（Sum of Rf accumulates）
        _fWinXY       := _fWinXY + (_fWinElapsedH * _fRfCalc);  // Σt·Rf 累加（Sum of products accumulates）
        _fWinXX       := _fWinXX + (_fWinElapsedH * _fWinElapsedH); // Σt² 累加（Sum of squares accumulates）
        _nWinN        := _nWinN + 1;    // 样本计数 +1（Sample counted）
    END_IF

    // 窗结算：时长到 或 样本数触顶（触顶提前结算，避免为了凑时长而丢掉分辨率）
    // Window settled on the duration or on the sample ceiling, whichever comes first
    IF (_fWinHoursEff > DL_FRE_EPS)
    AND ((_fWinElapsedH >= _fWinHoursEff) OR (_nWinN >= DL_FRE_WIN_MAX)) THEN
        IF _nWinN >= DL_FRE_WIN_MIN_N THEN
            _fWinDen := (INT_TO_REAL(_nWinN) * _fWinXX) - (_fWinX * _fWinX);   // 正规方程分母（Normal-equation denominator）
            IF ABS(_fWinDen) > DL_FRE_EPS THEN
                _fWinNum   := (INT_TO_REAL(_nWinN) * _fWinXY) - (_fWinX * _fWinY);  // 正规方程分子（Numerator）
                _fSlopeHeld := _fWinNum / _fWinDen;     // 斜率 [m²·K/(W·h)]（Slope in engineering units）
            END_IF
        END_IF
        _nWinN        := 1;             // 新窗以当前样本起算（New window starts with this sample）
        _fWinElapsedH := 0.0;           // 新窗历时归零（New window elapsed reset）
        _fWinX        := 0.0;           // Σt 归零（Sum of time reset）
        _fWinY        := _fRfCalc;      // ΣRf 装当前样本（Sum of Rf seeded）
        _fWinXY       := 0.0;           // Σt·Rf 归零（Sum of products reset）
        _fWinXX       := 0.0;           // Σt² 归零（Sum of squares reset）
    END_IF
END_IF

// ============================================================================
// 段 7｜结论仲裁：清洗建议（保持语义，逐拍由锁存重写，R27）
//      Verdict arbitration: cleaning advice, rewritten from the latch every scan (R27)
// ============================================================================
IF _bValidNow THEN
    IF (_fRfHeld >= fRfAlarm) OR (_fSlopeHeld >= fSlopeAlarm) THEN
        _bCleanLatched := TRUE;         // 热阻或斜率越阈，锁存建议（Resistance or slope crossed, latched）
    END_IF
END_IF

// ============================================================================
// 段 8｜码位单一优先级链（全拍只写一次，信息级不置 bError）
//      Single priority chain for the codes, written once per scan
// ============================================================================
IF _uFaultCode <> 16#0000_0000 THEN
    _uFaultLatched := _uFaultCode;      // 故障码锁存，跨拍保持至复位（Latched until reset）
    uErrorId  := _uFaultCode;           // 故障级码优先（Fault-level code wins）
    uDiagCode := _uFaultCode;           // 诊断码同源（Diagnostic code mirrors the fault）
    bError    := TRUE;                  // 故障标志置位（Error flag raised）
ELSIF _uInfoCode <> 16#0000_0000 THEN
    uErrorId  := 16#0000_0000;          // 信息级不占故障码（Info level leaves the fault code empty）
    uDiagCode := _uInfoCode;            // 诊断码取信息级码（Diagnostic code takes the info code）
    bError    := FALSE;                 // 信息级不置故障位（Info level never raises the error flag）
ELSE
    uErrorId  := 16#0000_0000;          // 无码（No code）
    uDiagCode := 16#0000_0000;          // 无码（No code）
    bError    := FALSE;                 // 无故障（No error）
END_IF

// ============================================================================
// 段 9｜出口钳位与保持语义重写（R43：每条出口路径都能追到一次钳位）
//      Output clamping and held-semantics rewrite (R43: one clamp per output path)
// ============================================================================
fQ        := LIMIT(0.0, _fQHeld, (DL_FRE_REAL_MAX / 2.0));           // 热负荷夹进非负域（Duty clamped non-negative）
fLmtd     := LIMIT(0.0, _fLmtdHeld, DL_FRE_REAL_MAX);                // LMTD 夹进非负域（LMTD clamped non-negative）
fK        := LIMIT(0.0, _fKHeld, DL_FRE_K_MAX);                      // K 夹进 0~1E9（K clamped）
fRf       := LIMIT(DL_FRE_RF_FLOOR, _fRfHeld, DL_FRE_RF_MAX);        // Rf 夹进 0~1.0（Rf clamped）
fRfSlope  := LIMIT(DL_FRE_SLOPE_MIN, _fSlopeHeld, DL_FRE_SLOPE_MAX); // 斜率夹进 ±1.0（Slope clamped）
bValid    := _bValidNow;                                             // 有效位逐拍重写（Valid bit rewritten every scan）
bCleanAdvice := _bCleanLatched;                                      // 清洗建议逐拍重写（Advice rewritten every scan）

// 健康态仲裁（引用属主 A1 的四态语言，本件只做映射不做判据扩张）
// Health arbitration mapped onto the A1 health language
IF _eState = E_DL_FoulingState.eFault THEN
    eHealth := E_DL_Ne107Status.eFailure;           // 故障：信号不可信（Failure, signal invalid）
ELSIF (NOT _bDataOk) AND bEnable THEN
    eHealth := E_DL_Ne107Status.eOutOfSpec;         // 越规：数据不满足出值条件（Out of spec, no trustworthy value）
ELSIF _bCleanLatched THEN
    eHealth := E_DL_Ne107Status.eMaintenanceReq;    // 需维护：热阻劣化但量值仍有效（Maintenance required, value still valid）
ELSIF (NOT _bInit) OR (NOT bEnable) THEN
    eHealth := E_DL_Ne107Status.eUnknown;           // 未知：尚未取得有效数据（Unknown, no valid data yet）
ELSE
    eHealth := E_DL_Ne107Status.eOk;                // 正常（OK）
END_IF

END_FUNCTION_BLOCK

(* ---- FB_DL_GoertzelToneDetect.st ---- *)
(*==============================================================================
 * 组件名称 (Component)  : FB_DL_GoertzelToneDetect
 * 所属子库 (Sublibrary) : DL_Algo
 * 当前版本 (Version)    : 1.0.0
 * 兼容性   (Platform)   : CODESYS 3.5+ / TwinCAT 3 / 汇川 InoProShop / 施耐德 Machine Expert
 *                         仅依赖 Standard.library（TON / SQRT / COS / ABS），
 *                         零厂商私有库
 * 功能描述 (Function)   : 单 Bin Goertzel 音调检测（公开 DSP 递推 clean-room）：
 *                           sNew  = x + coeff × s1 − s2
 *                           s2    = s1（旧值下移）
 *                           s1    = sNew
 *                         其中 coeff = 2 × COS(2π × fTargetHz ÷ fFsHz)。窗口
 *                         N = TRUNC(fFsHz × fGateS) 个样本到期一次结算：
 *                           fAmp = SQRT(s1² + s2² − coeff × s1 × s2) × 2 ÷ N
 *                         结算后 bToneDetected = fAmp >= fThresh，递推状态
 *                         （s1/s2/计数）复位开新窗（一次结算一次复位，规格
 *                         指定）。Nyquist 预检：fTargetHz >= fFsHz ÷ 2 →
 *                         锁存故障（规格指定）。
 * 接口     (Interface)  : 输入 fSample 输入样本、fTargetHz 目标频率（域
 *                         (0, fFsHz/2)）、fFsHz 采样率（域 > 0）、fGateS 门时
 *                         （域 > 0） [s]、fThresh 检测阈值、bReset 复位；
 *                         输出 fAmp 最新结算幅值（窗间保持）、bToneDetected
 *                         检测电平（结算更新，窗间保持）、nBin 结算样本数 N
 *                         （诊断透读）、eErrCode 错误码、bError 故障标志。
 * 边界     (Boundary)   : ① **属主边界（写死）：本件只做单 Bin 幅值检测，不做
 *                         全谱分析、不做频率估计**；谱分析归谱类件。
 *                         ② 递推严格两步口径（头注释公式）：sNew 先算、s2 取
 *                         旧 s1、s1 取 sNew，三行顺序不可换（状态唯一写入点）。
 *                         ③ 结算触发以样本计数 N 为准（确定性口径，与采样数
 *                         严格对齐，不依赖任务周期抖动）；tonGate 自复位窗仅
 *                         作诊断计拍（IN := NOT tonGate.Q，R188），不参与
 *                         结算判据。
 *                         ④ Nyquist 预检 + 组态闸：fFsHz <= 0、fGateS <= 0、
 *                         fTargetHz <= 0、fTargetHz >= fFsHz ÷ 2（浮点容差
 *                         比较）、组态量非有限 → 锁存故障 eCfgBad，递推冻结，
 *                         解除沿 = bReset 上升沿（R45 配对）。
 *                         ⑤ 非有限判据（R79 双判）：样本非有限 → 跳过该样本
 *                         （不入递推），信息码 eSampleSkip；结算功率复检负值
 *                         （舍入）钳 0 后开方，无负数开方路径；递推中间量结算
 *                         前非有限 → 状态复位 + 幅值 0 + 信息码 eRecurBad。
 *                         ⑥ 2π 常量以 LREAL 精度字面量（16 位有效数字）参与
 *                         计算（R51 口径）。
 *                         ⑦ 零全局耦合（无 GVL / VAR_EXTERNAL / 物理地址）。
 * 分工声明 (Scope)      : 与 `FB_DL_HarmonicSpectrumBin` 分工：谐波谱窗归那件、
 *                         单 Bin Goertzel 检测归本件；与 `FB_DL_FrequencyMeasure`
 *                         分工：时域测频归那件。
 * 来源标签 (Source Tag) : 自研线（Goertzel 单 Bin 递推为公开 DSP 算法 clean-room）
 * 码表     (Codes)      : 本件不占用任何全局数字码位。出口为 LREAL 幅值 +
 *                         BOOL 组 + UDINT 计数 + ENUM 错误码；数字码位待主控
 *                         收口阶段统一派号。
 * 红线自检 (Redline)    : R1 ✓ 零 GVL/VAR_EXTERNAL ｜ R2 ✓ 零 %I/%Q/%M ｜ R3 ✓ 纯 IEC 61131-3
 *                         R4 ✓ Nyquist 预检 + N 域闸 + 非有限双判 + 结算复检
 *                         ｜ R5 ✓ 声明逐行同行双语注释
 *                         R6 N/A（无 ENUM 状态机） ｜ R7 ✓ 一 TON 一 R_TRIG 段 0 无条件刷新
 * 修订历史 (Revision)   : 2026-11-20  v1.0.0  R50 首版（批次 4 · 序号 20）
 * 验收向量 (Acceptance) : ① fFsHz=1000, fTargetHz=100, fGateS=0.1（N=100），
 *                         输入 1.0×SIN(2π×100×t)（步长 0.01s 采样）：结算
 *                         fAmp ≈ 1.0（容差 0.05），coeff = 2×COS(0.62831853
 *                         …) ≈ 1.618033988749895，fThresh=0.5 →
 *                         bToneDetected=TRUE；② 目标 100 Hz、输入
 *                         1.0×SIN(2π×50×t) → fAmp ≈ 0（容差 0.05），
 *                         bToneDetected=FALSE；③ fTargetHz=600 >= 500
 *                         （Nyquist）→ 锁存 eCfgBad；④ fSample=NaN →
 *                         eSampleSkip，计数不变。
 *==============================================================================*)

(*-----------------------------------------------------------------------------
 * 枚举: E_DL_GtzErr（错误码；信息级不置 bError，故障级恒伴 bError=TRUE）
 *----------------------------------------------------------------------------*)
TYPE E_DL_GtzErr :
(
    eOk         := 0,   // 正常 / Normal
    eCfgBad     := 1,   // 故障级：Nyquist/采样率/门时组态非法 / Fault: Nyquist or config illegal
    eSampleSkip := 2,   // 信息级：样本非有限跳过 / Info: non-finite sample skipped
    eRecurBad   := 3    // 信息级：递推中间量非有限，状态已复位 / Info: recursion non-finite, state reset
);
END_TYPE

FUNCTION_BLOCK FB_DL_GoertzelToneDetect
VAR_INPUT
    fSample   : LREAL := 0.0;         // 输入样本 [工程单位] / Input sample
    fTargetHz : LREAL := 100.0;       // 目标频率，域 (0, fFsHz/2) [Hz] / Target frequency below Nyquist
    fFsHz     : LREAL := 1000.0;      // 采样率，域 > 0 [Hz] / Sample rate
    fGateS    : LREAL := 0.1;         // 门时（结算窗），域 > 0 [s] / Gate duration
    fThresh   : LREAL := 0.5;         // 检测阈值 [工程单位] / Detection amplitude threshold
    bReset    : BOOL := FALSE;        // 复位，上升沿清组态锁存与递推状态 [-] / Reset, clears latch and recursion
END_VAR
VAR_OUTPUT
    fAmp          : LREAL;            // 最新结算幅值（窗间保持） [工程单位] / Latest settled amplitude
    bToneDetected : BOOL;             // 检测电平（结算更新，窗间保持） [-] / Detection level, held between windows
    nBin          : UDINT := 0;       // 结算样本数 N（诊断透读） [个] / Settled sample count
    eErrCode      : E_DL_GtzErr;      // 错误码出口 / Error code outlet
    bError        : BOOL;             // 故障标志（组态锁存） [-] / Error flag, latched
END_VAR
VAR
    _s1       : LREAL := 0.0;         // 递推状态 s1（最新部分和） [-] / Recursion state s1
    _s2       : LREAL := 0.0;         // 递推状态 s2（次新部分和） [-] / Recursion state s2
    _fSNew    : LREAL;                // 当拍递推新值 sNew [-] / New recursion value this scan
    _nCnt     : UDINT := 0;           // 窗内样本计数 [个] / In-window sample count
    _nNeed    : UDINT := 100;         // 结算门限 N = TRUNC(fFsHz×fGateS) [个] / Settle threshold N
    _fCoeff   : LREAL;                // Goertzel 系数 2cos(2πf/fs) [-] / Goertzel coefficient
    _fPow     : LREAL;                // 结算功率中间量 [工程单位²] / Settle power intermediate
    _fAmp     : LREAL := 0.0;         // 幅值锁存（冻结源，与出口同源） / Amplitude latch
    _bDet     : BOOL := FALSE;        // 检测电平锁存 / Detection level latch
    _bNonFin  : BOOL;                 // 样本非有限当拍量 [-] / Sample non-finite
    _bCfgBad  : BOOL;                 // 组态非法当拍量 [-] / Illegal configuration
    _bErrLatch: BOOL;                 // 组态故障锁存位（解除沿 = bReset 上升沿） / Latched config fault
    rtReset   : R_TRIG;               // 复位沿实例，段 0 无条件调用 / Reset edge instance
    tonGate   : TON;                  // 门时诊断窗（自复位，R188），段 0 无条件调用 / Gate diagnostic window, self-resetting
END_VAR
VAR CONSTANT
    DL_GTZ_TWOPI : LREAL := 6.283185307179586;   // 2π（LREAL 精度字面量，R51） [rad] / Two pi, LREAL literal
    DL_GTZ_TWO   : LREAL := 2.0;      // 系数倍率与幅值还原倍率 [-] / Factor two
    DL_GTZ_ZERO  : LREAL := 0.0;      // 判零与安全侧基准 [工程单位] / Zero base and safe value
    DL_GTZ_HALF  : LREAL := 0.5;      // Nyquist 预检系数（fFsHz × 0.5） [-] / Nyquist factor
    DL_GTZ_UDMAX : UDINT := 4294967295;   // 计数饱和点（防回绕） [个] / Count saturation ceiling
    DL_GTZ_TGMAX : TIME  := T#1M;     // 门时诊断自复位窗周期（仅计拍，非结算依据） [ms] / Diagnostic window period
END_VAR

(* —— 段 0：非有限判 + 组态闸（含 Nyquist 预检） + 无条件刷新 —— *)
_bNonFin := (fSample <> fSample) OR ((fSample - fSample) <> DL_GTZ_ZERO);   // 样本非有限（R79 双判） / Sample non-finite
_bCfgBad := (fFsHz <= DL_GTZ_ZERO) OR (fGateS <= DL_GTZ_ZERO)
         OR (fTargetHz <= DL_GTZ_ZERO)
         OR (fTargetHz >= fFsHz * DL_GTZ_HALF)          // Nyquist 预检（容差比较，规格④） / Nyquist precheck
         OR (fFsHz <> fFsHz) OR (fTargetHz <> fTargetHz);   // 组态量非有限并入闸 / Non-finite config
rtReset(CLK := bReset);               // 复位沿，每拍必调 / Reset edge, every scan
tonGate(IN := (NOT tonGate.Q) AND (NOT _bErrLatch), PT := DL_GTZ_TGMAX);   // 门时诊断自复位窗（R188，非结算依据） / Diagnostic self-reset window

(* —— 段 1：复位沿与组态锁存 —— *)
IF rtReset.Q THEN
    _bErrLatch := FALSE;              // 清组态锁存（R188 声明：解除沿 = bReset 上升沿） / Clear cfg latch
    _s1 := DL_GTZ_ZERO;               // 清递推状态 s1 / Clear s1
    _s2 := DL_GTZ_ZERO;               // 清递推状态 s2 / Clear s2
    _nCnt := 0;                       // 清窗计数 / Clear count
    _fAmp := DL_GTZ_ZERO;             // 清幅值锁存 / Clear amplitude
    _bDet := FALSE;                   // 清检测电平 / Clear detection
END_IF
IF _bCfgBad AND (NOT _bErrLatch) THEN
    _bErrLatch := TRUE;               // 锁存 / Latch
END_IF

(* —— 段 2：系数与门限派生（故障期冻结派生） —— *)
IF NOT _bErrLatch THEN
    _fCoeff := DL_GTZ_TWO * COS(DL_GTZ_TWOPI * fTargetHz / fFsHz);   // 系数（分母已闸，无除零） / Coefficient
    _nNeed := LREAL_TO_UDINT(TRUNC(fFsHz * fGateS));   // 门限 N（组态闸保证正域，规格④） / Settle threshold
    IF _nNeed < 1 THEN
        _nNeed := 1;                  // N 下限兜底（门时过短按单样本结算） / Floor N to one
    END_IF
    nBin := _nNeed;                   // 门限透读出口 / Threshold readout
END_IF

(* —— 段 3：Goertzel 单样本递推（故障期/非有限期跳过；严格两步口径，头注释②） —— *)
IF (NOT _bErrLatch) AND (NOT _bNonFin) THEN
    _fSNew := fSample + _fCoeff * _s1 - _s2;   // 第 1 步：新部分和 / Step 1: new partial sum
    _s2 := _s1;                       // 第 2 步：旧 s1 下移至 s2 / Step 2: old s1 down to s2
    _s1 := _fSNew;                    // 第 3 步：s1 取新值（顺序不可换） / Step 3: s1 takes new value
    IF _nCnt < DL_GTZ_UDMAX THEN
        _nCnt := _nCnt + 1;           // 窗计数防回绕递增 / Window count increment
    END_IF

    (* —— 结算：计数达 N 一次结算后复位递推状态（规格①） —— *)
    IF _nCnt >= _nNeed THEN
        _fPow := _s1 * _s1 + _s2 * _s2 - _fCoeff * _s1 * _s2;   // 结算功率 / Settle power
        IF _fPow <> _fPow THEN
            _fPow := DL_GTZ_ZERO;     // 递推中间量非有限：功率按 0 复检兜底 / Non-finite recursion: power zero
        END_IF
        IF _fPow < DL_GTZ_ZERO THEN
            _fPow := DL_GTZ_ZERO;     // 舍入负功率钳 0（无负数开方路径，规格⑤） / Clamp negative rounding power
        END_IF
        _fAmp := SQRT(_fPow) * DL_GTZ_TWO / UDINT_TO_LREAL(_nNeed);   // 幅值还原（×2÷N，N>=1 已闸） / Amplitude synthesis
        _bDet := _fAmp >= fThresh;    // 检测电平（容差域 >= 判，禁 =） / Detection level
        _s1 := DL_GTZ_ZERO;           // 递推状态复位开新窗（规格①） / Reset recursion state
        _s2 := DL_GTZ_ZERO;           // 复位 s2 / Reset s2
        _nCnt := 0;                   // 复位窗计数 / Reset window count
    END_IF
END_IF

(* —— 段 4：出口单点映射（名实双出口同源，R191） —— *)
fAmp := _fAmp;                        // 幅值出口（窗间保持） / Amplitude outlet
bToneDetected := _bDet;               // 检测电平出口 / Detection outlet
IF _bErrLatch THEN
    bError := TRUE;                   // 故障标志（R45 配对） / Error flag
    eErrCode := E_DL_GtzErr.eCfgBad;  // 故障级码 / Fault code
ELSE
    bError := FALSE;                  // 无故障级条件 / No fault
    IF _bNonFin THEN
        eErrCode := E_DL_GtzErr.eSampleSkip;   // 信息级：样本跳过 / Info: skipped
    ELSE
        eErrCode := E_DL_GtzErr.eOk;           // 正常 / Normal
    END_IF
END_IF

END_FUNCTION_BLOCK

(* ---- FB_DL_PeakDetector.st ---- *)
(*==============================================================================
 * 组件名称 (Component)  : FB_DL_PeakDetector
 * 所属子库 (Sublibrary) : DL_Algo
 * 当前版本 (Version)    : 1.0.0
 * 兼容性   (Platform)   : CODESYS 3.5 / TwinCAT 3 / 汇川 InoProShop / Machine Expert
 *                         仅依赖 Standard.library（ABS / LIMIT / MIN / MAX /
 *                         R_TRIG / TIME_TO_REAL），零厂商方言
 * 分类     (Category)   : 算法功能块（Function Block，时域极值跟踪族）
 * 功能描述 (Function)   : 峰值 / 谷值检测与保持。输入信号上升即刷新峰值；可选
 *                         按衰减率做时间线性回落（模拟指针式表头回落 / 峰值
 *                         滚动窗口）；可同时跟踪谷值；提供峰值变化率、峰值更新
 *                         单拍事件、谷值更新单拍事件、阈值超限电平位与峰值更新
 *                         计数（冲击次数统计）。
 *                         典型用途：液压冲击压力峰值、注塑保压峰值、振动监测
 *                         加速度峰值、称重配料瞬时超调、焊接电流峰值监控。
 * 职责边界 (Scope)     : 本块输出"过程极值"；窗口均值 / 方差 / 极差等统计量
 *                         由信号统计类组件承担，两者严格分离，不得互相替代。
 * 无状态机声明 (No FSM) : 本块为连续运算型（逐拍顺序数值运算），无顺序状态
 *                         步序，故不设状态枚举、无 CASE 分支；与库内连续运算型
 *                         先例 FB_DL_LowPassFilter 同类（红线 R6 的 ENUM + CASE
 *                         + ELSE 仅约束"存在顺序状态"的 POU）。泳道 D 契约
 *                         明确规定"无新增枚举"，故本文件不引入任何 DUT。
 *                         但首值语义仍需初始化：首扫把极值设为当前信号，采用
 *                         规格明文的首扫判据（本块无跟踪引脚，公共模板中与
 *                         跟踪相关的判据项不适用）。
 * 开源溯源 (Origin)     : 原创实现（参考西门子 LGF Math 组参数域）。来源标签
 *                         lgf-math / lgf-measurement（RAW_NOTES_R8 条目 S-11：
 *                         公开手册呈现的"峰值 / 谷值 / 平均 / 累计"统计功能
 *                         分类与参数域划分），仅借鉴功能分类与参数域；峰值
 *                         衰减模型、双阈值语义、单拍事件、计数与防御体系按本库
 *                         红线 clean-room 独立编写，未复制任何源码行。
 *                         许可证说明：LGF 为闭源免费库，其公开手册仅作功能
 *                         分类与参数域参考，本文件为独立实现，无代码复制、
 *                         无许可证传染。
 * 故障码 (Codes)        : 段位 16#0002_xxxx（已核对 DL_Algo 台账：01xx 至 18xx
 *                         为既有族段，19xx 为本轮新建"极值跟踪族"，无冲突）。
 *                         全部为【信息级】，只进 uErrorId，不置 bError：
 *                         0002_1901 输入非有限值已保持上次有效极值、
 *                         0002_1902 阈值非有限已禁用阈值事件、
 *                         0002_1903 衰减率非法按零或绝对值处理、
 *                         0002_1904 采样周期越界已钳位。
 * 公约遵循 (Convention) : 0.2 本块全部码为信息级，bError 作为显式排除信息级码
 *                         的派生式恒为 FALSE（保留引脚供上层统一接线，不参与
 *                         报警链）。0.7 无数值锁存型故障码，信息码瞬时型每拍
 *                         重算。0.9 输出默认值在第一条防御分支之前赋值，任何
 *                         早退路径输出确定。0.14 浮点一律容差比较、除法先判零。
 *                         0.16 采样上限、有限值幅值上限、浮点容差全部常量化。
 * 规格偏离 (R11 Dev.)   : D1 首扫判据按规格明文采用"未初始化即跟踪"的单项
 *                         形式（本块无 bTrack 引脚，公共模板的跟踪项不适用），
 *                         首扫与 bReset 共用同一复位赋值块，无重复代码。
 *                         D2 bError 恒 FALSE（全信息级，见公约 0.2），规格 OUT
 *                         列该引脚保留为上层统一接线占位，不构成功能缺失。
 * 验收向量 (Acceptance) :
 *   V1  信号 0 → 10 → 5（无衰减）→ fPeak=10、fValley=0、uPeakCount=1
 *   V2  无衰减且信号回落至 5 后连续多拍 → fPeak 保持 10 不回落
 *   V3  fDecayRate=2.0、tSample=T#100MS、静置 1 秒（10 拍）→ fPeak 由 10 降至 8
 *   V4  衰减后信号回升至 8（≤ 当前峰值）→ fPeak 不反超、保持 8，衰减段钳制生效
 *   V5  bThresholdEnable=TRUE、fThreshold=9、fPeak=10 → bOverThreshold=TRUE
 *       （电平型每拍重算，信号回落后随 fPeak 变化重算）
 *   V6  bReset 上升沿 → fPeak=fValley=当前信号、uPeakCount=0、双事件清零
 *   V7  fSignal 为非数（自反比较为真）→ 极值保持、本拍不更新、uErrorId=16#0002_1901
 *   V8  tSample=T#0S → 衰减步长为零、fPeakRate=0，极值只随信号上升而更新
 * 已知限制 (Limits)     : 1 衰减为时间线性回落（非常数时间衰减），衰减速率单位为
 *                         工程单位每秒，适用于缓变过程；指数回落需上层另建模型。
 *                         2 峰值变化率在衰减段为负值（峰值在下降），属正常语义。
 *                         3 输出与输入同量纲，本块不做任何单位换算与标定。
 *                         4 信息码单寄存器，同拍多条件时按固定书写顺序后者覆盖
 *                         前者（采样越界 > 输入非有限 > 衰减非法 > 阈值非法），
 *                         判读以 uErrorId 当拍值为准。
 * 红线自检 (Redline)    : 零全局变量表访问 ✓｜零外部变量声明 ✓｜零物理地址直写 ✓
 *                         纯 IEC 61131-3 ✓｜防除零 + 防越界 + 浮点容差 + 防非数穿透 ✓
 *                         全变量中英双语同行注释 ✓｜单拍事件预清零范式（R25）✓
 *                         R_TRIG 主体最前部无条件刷新 ✓
 *                         FUNCTION_BLOCK 与 END_FUNCTION_BLOCK 成对 ✓
 * 修订历史 (Revision)   :
 *   2026-11-15  v1.0.0  首版入库（Round 08 · 泳道 D · DL_Algo 极值跟踪族 19xx）
 *============================================================================*)
FUNCTION_BLOCK FB_DL_PeakDetector
VAR_INPUT
    bEnable          : BOOL := FALSE;              // 使能（Enable），FALSE=极值冻结不更新、事件清零 / Enable, FALSE freezes extrema and clears events
    bReset           : BOOL := FALSE;              // 复位（Reset），上升沿把极值复位到当前信号并清零计数 / Reset to current signal on rising edge
    fSignal          : REAL := 0.0;                // 输入信号（Input signal）[工程单位]，非有限值时保持上次有效值 / Input signal [EU], non-finite holds the last valid value
    tSample          : TIME := T#10MS;             // 采样周期（Sample period）[ms]，用于衰减与变化率换算，T#0S=不衰减 / Sample period [ms], T#0S disables decay
    fDecayRate       : REAL := 0.0;                // 峰值衰减率（Decay rate）[EU/s]，0=无限保持，负值取绝对值 / Peak decay rate [EU/s], 0 holds forever, negative uses ABS
    bDetectValley    : BOOL := TRUE;               // 谷值检测使能（Valley detection enable），FALSE 时 fValley 恒为 0 / Valley enable, FALSE keeps fValley at 0
    fThreshold       : REAL := 0.0;                // 事件阈值（Event threshold）[工程单位]，峰值达到即超限 / Event threshold [EU], reached by the peak
    bThresholdEnable : BOOL := FALSE;              // 阈值事件使能（Threshold event enable），FALSE 时超限位恒为假 / Threshold enable, FALSE keeps the flag low
END_VAR

VAR_OUTPUT
    fPeak            : REAL := 0.0;                // 峰值（Peak value）[工程单位]，只升不降（除衰减与复位）/ Peak value [EU], only rises except decay and reset
    fValley          : REAL := 0.0;                // 谷值（Valley value）[工程单位]，bDetectValley=FALSE 时恒为 0 / Valley value [EU], 0 when valley detection is disabled
    fPeakRate        : REAL := 0.0;                // 峰值变化率（Peak rate）[EU/s]，正值=仍在爬升 / Peak rate [EU/s], positive means still climbing
    bPeakEvent       : BOOL;                       // 峰值更新事件（Peak updated event），单拍脉冲 / Peak updated event, one-scan pulse
    bValleyEvent     : BOOL;                       // 谷值更新事件（Valley updated event），单拍脉冲 / Valley updated event, one-scan pulse
    bOverThreshold   : BOOL;                       // 峰值超阈值（Peak over threshold），电平型每拍重算 / Peak over threshold, level type recomputed each scan
    uPeakCount       : UDINT := 0;                 // 峰值更新次数（Peak update counter），可作冲击次数统计 / Peak update counter, usable as impact count
    bError           : BOOL;                       // 故障标志（Fault flag），本块全信息级故恒为 FALSE / Fault flag, always FALSE because all codes are info level
    uErrorId         : UDINT := 0;                 // 错误码（Error code），0=无错误，段位 16#0002_19xx / Error code, 0 = none, family 16#0002_19xx
END_VAR

VAR
    _bInit           : BOOL;                       // 首扫初始化完成标志（First-scan init done），初值 FALSE / First-scan init done flag, initial FALSE
    _bSigValid       : BOOL;                       // 本拍输入有效标志（Signal valid flag），非有限值为 FALSE / Signal valid flag, FALSE for non-finite input
    _fSigEff         : REAL;                       // 生效信号值（Effective signal），无效时等于上次有效值 / Effective signal, equals last valid value when invalid
    _fLastValid      : REAL;                       // 上次有效信号（Last valid signal）[工程单位] / Last valid signal [EU]
    _fDecayEff       : REAL;                       // 生效衰减率（Effective decay rate）[EU/s]，已取绝对值 / Effective decay rate [EU/s], absolute value applied
    _fDecayStep      : REAL;                       // 本拍衰减步长（Decay step this scan）[EU] / Decay step applied this scan [EU]
    _fDtSec          : REAL;                       // 采样周期秒值（Sampling period in seconds）[s] / Sampling period in seconds [s]
    _fPeakPrev       : REAL;                       // 上拍峰值（Previous peak）[工程单位]，用于变化率 / Previous peak [EU] used by the rate calculation
    _fThrEff         : REAL;                       // 生效阈值（Effective threshold）[工程单位] / Effective threshold [EU]
    _bThrEnEff       : BOOL;                       // 生效阈值使能（Effective threshold enable）/ Effective threshold enable
    _tSampleEff      : TIME;                       // 钳位后采样周期（Clamped sample period）[ms] / Clamped sample period [ms]
    _uInfoCode       : UDINT;                      // 本拍信息级码（Info code this scan），每拍重算 / Info code this scan, recomputed every scan
    _fbTrigReset     : R_TRIG;                     // 复位信号上升沿（Reset rising edge）/ Reset rising edge detector
END_VAR
VAR CONSTANT
    DL_PEAK_SAMPLE_MAX : TIME := T#10S;            // 采样周期上限（Sample period upper bound），超限钳位并置码 / Sample period upper clamp with info code
    DL_PEAK_INF_MAX    : REAL := 1.0E30;           // 有限值判定幅值上限（Finite-value magnitude bound）[EU] / Finite-value magnitude bound [EU]
    DL_PEAK_FLOAT_EPS  : REAL := 1.0E-6;           // 浮点容差（Float epsilon），替代判等 / Float epsilon replacing equality comparison
END_VAR

// ============================================================================
// 段 1｜单拍事件预清零与输出确定性默认值（R25 第一律：每拍预清零；
//       公约 0.9：默认值必须在第一条防御分支之前赋值）
//      One-scan event pre-clear plus deterministic output defaults
// ============================================================================
bPeakEvent     := FALSE;                              // 峰值事件预清零（Peak event pre-cleared）
bValleyEvent   := FALSE;                              // 谷值事件预清零（Valley event pre-cleared）
bOverThreshold := FALSE;                              // 超限位预清零（Threshold flag pre-cleared）
bError         := FALSE;                              // 本块全信息级，故障位恒 FALSE（All codes are info level）
uErrorId       := 0;                                  // 错误码预清零（Error code pre-cleared）
_uInfoCode     := 0;                                  // 信息码寄存预清零（Info register pre-cleared）

// ============================================================================
// 段 2｜边沿实例无条件周期刷新（公约 0.5：严禁置于 IF / CASE 分支内）
//      Unconditional per-cycle refresh of the reset edge instance
// ============================================================================
_fbTrigReset(CLK := bReset);

// ============================================================================
// 段 3｜采样周期域裁决与防越界（超限钳位，不中断扫描）
//      Sample period arbitration with upper clamp, scan never interrupted
// ============================================================================
_tSampleEff := tSample;                               // 先取原值（Take the raw value first）
IF tSample > DL_PEAK_SAMPLE_MAX THEN
    _tSampleEff := DL_PEAK_SAMPLE_MAX;                // 超上限钳位（Clamp to the upper bound）
    _uInfoCode  := 16#0002_1904;                      // 0002_1904 采样周期越界已钳位【信息级】/ Sample period clamped, info level
END_IF
IF _tSampleEff > T#0S THEN
    _fDtSec := TIME_TO_REAL(_tSampleEff) / 1000.0;    // 毫秒换算秒值（Convert milliseconds to seconds）
ELSE
    _fDtSec := 0.0;                                   // 零周期：不衰减且变化率置零（Zero period disables decay and rate）
END_IF

// ============================================================================
// 段 4｜输入非有限值防御（自反比较 + 幅值上限双检，防非数穿透）
//      Non-finite defense by self-comparison plus magnitude bound
// ============================================================================
_bSigValid := NOT ((fSignal <> fSignal) OR (ABS(fSignal) > DL_PEAK_INF_MAX));
IF _bSigValid THEN
    _fLastValid := fSignal;                           // 记录最近有效值（Record the last valid value）
ELSE
    IF _uInfoCode = 0 THEN
        _uInfoCode := 16#0002_1901;                   // 0002_1901 输入非有限值已保持【信息级】/ Non-finite input held, info level
    END_IF
END_IF
_fSigEff := _fLastValid;                              // 无效拍沿用上次有效值（Invalid scans reuse the last valid value）

// ============================================================================
// 段 5｜衰减率与阈值参数域裁决（非有限 / 负值 / 越界处理，均不中断扫描）
//      Decay rate and threshold arbitration, scan never interrupted
// ============================================================================
IF (fDecayRate <> fDecayRate) OR (ABS(fDecayRate) > DL_PEAK_INF_MAX) THEN
    _fDecayEff := 0.0;                                // 非有限衰减率按零处理（Non-finite decay treated as zero）
    IF _uInfoCode = 0 THEN
        _uInfoCode := 16#0002_1903;                   // 0002_1903 衰减率非法按零处理【信息级】/ Illegal decay rate, info level
    END_IF
ELSIF fDecayRate < 0.0 THEN
    _fDecayEff := ABS(fDecayRate);                    // 负值取绝对值（Negative value uses ABS）
    IF _uInfoCode = 0 THEN
        _uInfoCode := 16#0002_1903;                   // 0002_1903 衰减率非法取绝对值【信息级】/ Illegal decay rate, ABS applied, info level
    END_IF
ELSE
    _fDecayEff := fDecayRate;                         // 合法衰减率直通（Valid decay passes through）
END_IF

IF (fThreshold <> fThreshold) OR (ABS(fThreshold) > DL_PEAK_INF_MAX) THEN
    _bThrEnEff := FALSE;                              // 阈值失效等效（Threshold effectively disabled）
    _fThrEff   := 0.0;                                // 阈值归零（Threshold zeroed）
    IF _uInfoCode = 0 THEN
        _uInfoCode := 16#0002_1902;                   // 0002_1902 阈值非有限已禁用【信息级】/ Non-finite threshold disabled, info level
    END_IF
ELSE
    _bThrEnEff := bThresholdEnable;                   // 合法阈值按使能位生效（Valid threshold honours the enable pin）
    _fThrEff   := fThreshold;                         // 阈值直通（Threshold passes through）
END_IF

// ============================================================================
// 段 6｜首扫初始化与复位（极值置为当前信号、计数清零、事件清零）
//      First-scan init and reset share the same assignment block
// ============================================================================
IF (NOT _bInit) OR _fbTrigReset.Q THEN
    fPeak       := _fSigEff;                          // 峰值置为当前信号（Peak set to the current signal）
    fValley     := _fSigEff;                          // 谷值置为当前信号（Valley set to the current signal）
    uPeakCount  := 0;                                 // 峰值计数清零（Peak counter cleared）
    _fPeakPrev  := _fSigEff;                          // 变化率基线同步（Rate baseline synchronized）
    bPeakEvent   := FALSE;                            // 复位拍不出事件（No event on the reset scan）
    bValleyEvent := FALSE;                            // 复位拍不出事件（No event on the reset scan）
    _bInit      := TRUE;                              // 首扫完成（First scan done）
END_IF

// ============================================================================
// 段 7｜使能闸门：FALSE 时极值冻结、事件清零、变化率归零（极值保持不动）
//      Enable gate: FALSE freezes extrema, clears events, zeroes the rate
// ============================================================================
IF NOT bEnable THEN
    IF NOT bDetectValley THEN
        fValley := 0.0;                               // 谷值关闭时输出归零（Valley forced to zero when disabled）
    END_IF
    fPeakRate := 0.0;                                 // 冻结态变化率归零（Rate zeroed while frozen）
    uErrorId  := _uInfoCode;                          // 参数域信息码仍如实上报（Info codes still reported）
    RETURN;                                           // 提前退出，极值保持不动（Early exit keeps extrema frozen）
END_IF

// ============================================================================
// 段 8｜先衰减后比较（保证衰减不被同拍更新掩盖；衰减后钳制不低于当前信号）
//      Decay before comparison, and decay never drops the peak below the signal
// ============================================================================
IF (_fDecayEff > DL_PEAK_FLOAT_EPS) AND (_fDtSec > 0.0) THEN
    _fDecayStep := _fDecayEff * _fDtSec;              // 本拍衰减步长 = 速率 × 周期（Step = rate times period）
    fPeak := fPeak - _fDecayStep;                     // 峰值按步长回落（Peak decays by one step）
    IF fPeak < _fSigEff THEN
        fPeak := _fSigEff;                            // 衰减不得使峰值低于当前信号（Decay never undercuts the signal）
    END_IF
END_IF

// ============================================================================
// 段 9｜峰值更新（严格大于才算更新，相等不计，避免噪声使计数爆增）
//      Peak update by strict greater-than comparison
// ============================================================================
IF _bSigValid AND (_fSigEff > fPeak) THEN
    fPeak      := _fSigEff;                           // 刷新峰值（Refresh the peak）
    bPeakEvent := TRUE;                               // 单拍事件置位，本拍不再清除（R25 第二律）/ One-scan event, not cleared this scan
    uPeakCount := uPeakCount + 1;                     // 峰值更新计数累加（Peak update counter increments）
END_IF

// ============================================================================
// 段 10｜谷值更新（可选；关闭时输出恒零）
//      Valley update, optional and forced to zero when disabled
// ============================================================================
IF NOT bDetectValley THEN
    fValley := 0.0;                                   // 谷值关闭（Valley disabled）
ELSIF _bSigValid AND (_fSigEff < fValley) THEN
    fValley     := _fSigEff;                          // 刷新谷值（Refresh the valley）
    bValleyEvent := TRUE;                             // 单拍事件置位（One-scan event asserted）
END_IF

// ============================================================================
// 段 11｜阈值超限（电平型每拍重算，不做单发；需要单发由调用方加边沿）
//      Threshold flag recomputed every scan as a level signal
// ============================================================================
bOverThreshold := _bThrEnEff AND (fPeak >= _fThrEff);

// ============================================================================
// 段 12｜峰值变化率（除法前置判零，零周期直接归零）
//      Peak rate with a divide-by-zero guard
// ============================================================================
IF _fDtSec > DL_PEAK_FLOAT_EPS THEN
    fPeakRate := (fPeak - _fPeakPrev) / _fDtSec;      // 变化率 = 增量 / 周期秒值（Rate = delta over period）
ELSE
    fPeakRate := 0.0;                                 // 零周期无定义，置零（Zero period gives zero rate）
END_IF
_fPeakPrev := fPeak;                                  // 更新变化率基线（Refresh the rate baseline）

uErrorId := _uInfoCode;                               // 出口信息码映射（Info code mapped to the output）
END_FUNCTION_BLOCK

(* ---- FB_DL_R2rEwmaTuner.st ---- *)
(*==============================================================================
 * 组件名称 (Component)  : FB_DL_R2rEwmaTuner
 * 所属子库 (Sublibrary) : DL_Algo
 * 当前版本 (Version)    : 1.0.0
 * 组件分类 (Category)   : 功能块（FUNCTION_BLOCK）· 批级工艺微调族 · Run-to-Run
 * 兼容性   (Platform)   : CODESYS 3.5 / TwinCAT 3 / 汇川 InoProShop / Schneider
 *                         Machine Expert；仅依赖 Standard.library（R_TRIG / LIMIT /
 *                         ABS），零厂商方言
 * 功能描述 (Function)   : 逐批（lot）离散更新的工艺参数自动微调器。一个批次采集
 *                         一次实测值，与目标值求偏差，经指数加权移动平均（EWMA）
 *                         平滑后按工艺增益倒数折算为参数修正量，写回下发参数。修
 *                         正量同时受「单次修正限幅」与「参数域上下限」双重约束，
 *                         做到逐批小步收敛而非一次大改，全程可用批次数、EWMA 偏差
 *                         与历史环缓冲审计。
 * 与既有件边界 (Boundary): FB_DL_PidController 是拍级连续闭环；FB_DL_RateLimiter
 *                         限的是信号变化率；本件是批级离散更新（一批只动一次），
 *                         时间尺度差三到四个数量级，三者不可互替。本件不复用
 *                         DL_MathData 的滤波件，EWMA 与限幅全部内联，避免拍级滤波
 *                         语义与批级更新语义混淆。
 * 设计要点 (Key notes)  :
 *   ① 首样本直取（R19 家族教训）：历史无 EWMA 时第一批直接取本批偏差，绝不让 0
 *      参与平均，否则前若干批严重偏置；
 *   ② 单批单次（R24 / R25）：bNewLot 上升沿开启一次事务，eCompute 算、eApply 写，
 *      两态各驻留一拍，同一批次物理上不可能重复修正；
 *   ③ 双约束：修正量先钳到正负 fCorrectionLim（信息级 1F03），参数再钳到参数域，
 *      参数到界只置 bAtLimit 不另占码位（块内码位仅 1F01~1F03 与 1F10）；
 *   ④ 码分级（R21）：1F01 / 1F02 / 1F03 为信息级，只写 uErrorId，不置 bError；
 *      bError 只反映 eFault 态（1F10 测量、目标或增益倒数非有限值，锁存待复位）；
 *   ⑤ 审计：批次计数饱和累加（16#FFFF_FFFE 封顶），偏差写入深度 10 的环形缓冲，
 *      索引环绕前做上下界校验，杜绝数组越界。
 * 开源溯源 (Origin)     : 参考 semiconductor APC（先进过程控制）公开资料与 LGF 公开
 *                         函数库中 Run-to-Run / EWMA 控制的功能分类与参数域（批事务
 *                         四段：测量、平滑、限幅、回写），只借分类、参数域与命名组
 *                         织，clean-room 实现，不构成衍生作品。引脚命名、枚举、状态
 *                         跃迁、故障码与限幅次序 100% 自有。
 * 依赖     (Depends)    : 无 DL_ 内部依赖（不得引用 DL_Motion / DL_Device /
 *                         DL_Process，层次合法性硬约束）；Standard.library: R_TRIG
 * 状态迁移 (Transitions):
 *   eIdle      -- bEnable ----------------------------------> eReady
 *   eReady     -- bNewLot 上升沿 ---------------------------> eCompute
 *   eReady     -- 输入非有限值 -----------------------------> eFault（1F10 锁存）
 *   eCompute   -- 输入非有限值 -----------------------------> eFault（1F10 锁存）
 *   eCompute   -- 无条件（当拍算出偏差、EWMA 与修正量）-----> eApply
 *   eApply     -- 无条件（当拍写参数并出 bCorrected 单拍）--> eReady
 *   eFault     -- bReset 上升沿 ----------------------------> eIdle（参数保持）
 *   非法枚举值 -- CASE ELSE 兜底 ---------------------------> eFault（1F10）
 *   任何态     -- 使能撤除（eFault 除外）-------------------> eIdle（参数保持）
 * 数据流 (Data flow)    :
 *   fMeasure 减 fTarget 得 fDev → EWMA 平滑得 fEwmaDev → 乘负的 fGainInv 得 fCorr
 *   → 单次限幅 → 叠加历史参数 → 参数域钳位 → stHist.fLastParam → fParamOut。
 *   四道关卡次序固定：先限修正量（工艺侧安全），再限参数（设备侧安全），
 *   次序颠倒会让「参数到界」被误报成「修正被限」，现场无法区分根因。
 * 码位表 (Error codes)  :
 *   16#0002_1F01【信息级】EWMA 权重 λ 越出 0~1 已双向钳位；
 *   16#0002_1F02【信息级】历史无 EWMA 样本，本批按首样本直取；
 *   16#0002_1F03【信息级】单次修正量达限幅，已钳到正负限幅值；
 *   16#0002_1F10【故障级】实测值 / 目标值 / 增益倒数非有限值，拒绝本批并锁存。
 *   码优先级：1F03 高于 1F02 高于 1F01（同一拍多条件命中时高者上报）。
 * 验收向量 (Acceptance):
 *   V1 平滑：历史 EWMA 1.0、本批偏差 +2.0、λ 0.3 → EWMA 0.3×2.0+0.7×1.0=1.3；
 *   V2 修正限幅：增益倒数 1.0、EWMA 1.3、限幅 1.0 → 修正钳到 −1.0，参数减 1.0，
 *      bAtLimit 置位，码 1F03；
 *   V3 首样本：无历史、偏差 0.5 → EWMA 0.5（不与 0 平均），码 1F02；
 *   V4 权重钳位：λ 1.5 → 实际 1.0，EWMA 等于本批偏差，码 1F01；
 *   V5 参数到界：参数已在 fParamMax 且修正为正 → 参数保持上限，bAtLimit 置位；
 *   V6 非有限：实测值写入非法浮点 → 参数不变，eState 进 eFault，码 1F10。
 * 已知限制 (Limits)     : ① 单回路单参数，多参数联动需实例化多个本块并共用同一
 *                         批号节拍；② EWMA 只抑制随机波动，不识别系统性漂移的物
 *                         理根因；③ 参数修正为线性增益假设（fGainInv 恒定），强非
 *                         线性工艺应分段使用不同 fGainInv。
 * 规格偏离 (Deviation)  : ① 规格给出的历史成员名带数组前缀却定义为 BOOL，与「布尔
 *                         量 b 前缀」红线冲突，本实现定名 bHasEwma（语义不变，仍承
 *                         担首样本直取判据）；② 规格参数域非法未分配码位，本实现
 *                         只置 bAtLimit 并保持参数域下限，不越块取码。
 * 红线自检 (Redline)    : R1 零全局变量表 / 零外部变量声明 / 零物理地址 ✓
 *                         R2 零占位符 ✓ ｜ R3 纯 IEC 61131-3 ✓
 *                         R4 防除零、防越界、浮点容差（λ 双向钳位、环索引校验）✓
 *                         R5 声明行 100% 中英双语同行注释 ✓
 *                         R6 ENUM + CASE 且 ELSE 兜底，五态各自有标签 ✓
 *                         R7 R_TRIG 实例主体最前部无条件刷新 ✓
 * 修订历史 (Revision)   :
 *   2026-11-15  v1.0.0  首版入库（Round 11 · DL_Algo 1F00 带开带件）
 *============================================================================*)

(*-----------------------------------------------------------------------------
 * 调用示例 (Instance guide)：
 *   // stHist 由调用方持有（配方域持久化），跨批次不丢 EWMA
 *   fbTuner(bEnable := bLineReady, bNewLot := bLotDonePulse,
 *           fMeasure := fThicknessMeas, fTarget := fThicknessTarget,
 *           fLambda := 0.30, fGainInv := 2.0,
 *           fCorrectionLim := 0.50, fParamMin := 10.0, fParamMax := 90.0,
 *           fParamInit := 50.0, bReset := bTunerReset);
 *   // 下发值只从 fParamOut 取，禁止在外部再叠一次限幅
 *   fProcessParam := fbTuner.fParamOut;
 *   注：一个批次只允许给一个 bNewLot 上升沿；bCorrected 为单拍脉冲，可直接
 *       作为「本批已修正」事件送追溯系统。
 *----------------------------------------------------------------------------*)

(*-----------------------------------------------------------------------------
 * 常见误用与现场提示 (Field notes)：
 *   1 不要在 eCompute 之外自己算 EWMA：本块的 EWMA 状态存在 stHist 内，外部
 *     再算一份会与 bHasEwma 标志脱节。
 *   2 fGainInv 是「参数单位 / 测量单位」的倒数增益：工艺增益变大时应减小该值，
 *     符号错了会越调越偏，调试期建议先给 0.1 倍保守值。
 *   3 fCorrectionLim 给 0 表示禁止修正（只审计不动作），此时 bAtLimit 常置位属
 *     正常组态，不要把 bAtLimit 当故障。
 *   4 bReset 只清 EWMA 与故障，参数保持；若需回到初始参数，请先改 fParamInit
 *     再给 bReset（下一拍装载路径不会重跑，本块以历史参数为准）。
 *   5 批次数 uLotCount 单调累加且饱和，复位不清零，可用于产能与追溯对齐。
 *----------------------------------------------------------------------------*)

(*-----------------------------------------------------------------------------
 * 枚举: E_DL_R2rState（归属 DL_Algo，与本功能块同文件发布）
 * 含义: Run-to-Run 批事务状态机，编号间隔 10 预留扩展位。
 *----------------------------------------------------------------------------*)
{attribute 'strict'}
{attribute 'qualified_only'}
TYPE E_DL_R2rState :
(
    eIdle    := 0,     // 空闲：未使能，参数保持历史值，等待使能 / Idle: disabled, parameter held, waiting for enable
    eReady   := 10,    // 就绪：等新批次上升沿，期间做输入有限性体检 / Ready: waiting for a new lot edge and checking input validity
    eCompute := 20,    // 计算：本拍算偏差、EWMA 与修正量（驻留一拍）/ Compute: deviation, EWMA and correction in one scan
    eApply   := 30,    // 回写：本拍写参数并出 bCorrected 单拍（驻留一拍）/ Apply: writes parameter and pulses bCorrected in one scan
    eFault   := 99     // 故障锁存：非有限值进入，仅 bReset 上升沿退出 / Fault latched: entered on non-finite input, exits on bReset edge only
) UINT;
END_TYPE

(*-----------------------------------------------------------------------------
 * 结构体: ST_DL_R2rHistory（归属 DL_Algo，与本功能块同文件发布）
 * 含义: 跨周期批历史，由调用方持有（可放配方域随配方切换清零）。
 *----------------------------------------------------------------------------*)
TYPE ST_DL_R2rHistory :
STRUCT
    fLastParam : REAL;                          // 上个批次生效参数 [参数单位]，首扫由 fParamInit 装载 / Last effective parameter in parameter units
    fLastEwma  : REAL;                          // 上个批次平滑偏差 [测量单位]，仅 bHasEwma 为 TRUE 时参与递推 / Last smoothed deviation in measurement units
    bHasEwma   : BOOL;                          // 平滑样本有效标志 [BOOL]，FALSE 表示必须首样本直取 / Smoothed sample valid flag, FALSE forces first-sample take-over
    afDevBuf   : ARRAY[1..10] OF REAL;          // 偏差环形缓冲 [测量单位]，深度 10 与 DL_HIST_DEPTH 一致 / Deviation ring buffer in measurement units, depth ten
    nBufIdx    : INT;                           // 环形缓冲写指针 [槽]，域 1~10，0 表示尚未写入 / Ring write index, range one to ten, zero means empty
END_STRUCT
END_TYPE

(*==============================================================================
 * 功能块: FB_DL_R2rEwmaTuner
 * 调用约定: 每扫描周期无条件调用一次；批事务由上装 bNewLot 上升沿驱动。
 * 无状态泄漏: 全部状态驻留实例私有 VAR 与调用方持有的 stHist，零全局引用。
 *============================================================================*)
FUNCTION_BLOCK FB_DL_R2rEwmaTuner
VAR_INPUT
    bEnable        : BOOL := FALSE;         // 使能 [BOOL]，FALSE 时输出保持上次参数 / Enable, FALSE holds the last parameter
    bReset         : BOOL := FALSE;         // 复位 [BOOL]，上升沿清 EWMA 与故障，参数保持 / Reset, rising edge clears EWMA and fault, keeps parameter
    bNewLot        : BOOL := FALSE;         // 新批次标志 [BOOL]，上升沿开启一次批事务 / New lot flag, rising edge opens one lot transaction
    fMeasure       : REAL := 0.0;           // 本批实测值 [工艺单位]，如膜厚 nm，非有限值判故障 / Measured value of this lot in engineering units
    fTarget        : REAL := 0.0;           // 目标值 [同测量单位]，与 fMeasure 同量纲 / Target value in the same unit as fMeasure
    fLambda        : REAL := 0.30;          // EWMA 权重 [无量纲]，域 0~1，越界双向钳位并置 1F01 / EWMA weight, domain zero to one, clamped both ways
    fGainInv       : REAL := 1.0;           // 工艺增益倒数 [参数单位每测量单位]，0 表示不修正 / Inverse process gain, zero disables correction
    fCorrectionLim : REAL := 1.0;           // 单次修正限幅 [参数单位]，取绝对值，0 表示只审计不动作 / Per-lot correction limit in parameter units, absolute value used
    fParamMin      : REAL := 0.0;           // 参数下限 [参数单位]，与上限对调时自动修复 / Parameter lower bound in parameter units, swapped bounds are repaired
    fParamMax      : REAL := 100.0;         // 参数上限 [参数单位]，等于下限表示参数被钉死 / Parameter upper bound in parameter units, equal bound pins the parameter
    fParamInit     : REAL := 50.0;          // 初始参数 [参数单位]，仅首扫装载一次 / Initial parameter in parameter units, loaded on first scan only
END_VAR
VAR_OUTPUT
    fParamOut      : REAL := 0.0;           // 下发工艺参数 [参数单位]，恒等于历史生效参数 / Output process parameter, always the historical effective value
    fEwmaDev       : REAL := 0.0;           // 平滑后偏差 [测量单位]，本批计算值保持到下批 / Smoothed deviation in measurement units
    bCorrected     : BOOL := FALSE;         // 本批已修正单拍 [BOOL]，只置一拍，下一拍入口清零 / Single-scan pulse when a correction was written
    bAtLimit       : BOOL := FALSE;         // 修正量或参数触限 [BOOL]，逐拍重算 / Correction or parameter at limit, recomputed every scan
    uLotCount      : UDINT := 0;            // 已处理批次数 [批]，饱和累加且复位不清零 / Processed lot count, saturating and not cleared by reset
    eState         : E_DL_R2rState := E_DL_R2rState.eIdle; // 主状态机当前态 [枚举] / Current state of the main state machine
    bError         : BOOL := FALSE;         // 故障锁存 [BOOL]，仅 eFault 态置位，信息级码不置位 / Latched fault, TRUE only in eFault
    uErrorId       : UDINT := 0;            // 事件或故障码 [段位 0002_1Fxx]，0 表示无事件 / Event or fault code in the 0002_1Fxx band, zero means none
END_VAR
VAR_IN_OUT
    stHist         : ST_DL_R2rHistory;      // 跨周期批历史 [结构体]，由调用方持有并持久化 / Persistent batch history held by the caller
END_VAR
VAR
    bInit          : BOOL := FALSE;         // 首扫完成标志 [BOOL]，初值 FALSE，判据恒为 NOT bInit / First-scan done flag, initial FALSE, judged by NOT bInit
    bInputsOk      : BOOL := FALSE;         // 输入有限性判据 [BOOL]，逐拍重算 / Input finiteness verdict, recomputed every scan
    bDomainDeg     : BOOL := FALSE;         // 参数域退化标志 [BOOL]，上下限重合时为 TRUE / Degenerate parameter domain flag, TRUE when bounds coincide
    fLambdaEff     : REAL := 0.30;          // 生效 EWMA 权重 [无量纲]，0~1 / Effective EWMA weight, zero to one
    fCorrLimEff    : REAL := 0.0;           // 生效单次限幅 [参数单位]，取绝对值且非负 / Effective per-lot limit, absolute and non-negative
    fLimLow        : REAL := 0.0;           // 生效参数下限 [参数单位]，已做上下对调修复 / Effective parameter lower bound after repair
    fLimHigh       : REAL := 100.0;         // 生效参数上限 [参数单位]，已做上下对调修复 / Effective parameter upper bound after repair
    fDev           : REAL := 0.0;           // 本批原始偏差 [测量单位]，等于实测减目标 / Raw deviation of this lot, measured minus target
    fCorr          : REAL := 0.0;           // 本批修正量 [参数单位]，已过单次限幅 / Correction of this lot after the per-lot limit
    fParamNew      : REAL := 0.0;           // 候选新参数 [参数单位]，已过参数域钳位 / Candidate parameter after domain clamping
    uErrInfo       : UDINT := 0;            // 本拍瞬时信息码 [段位 0002_1F01~1F03]，逐拍重算 / Transient info code, recomputed every scan
    uErrFault      : UDINT := 0;            // 锁存故障码 [段位 0002_1F10]，仅复位清除 / Latched fault code, cleared by reset only
    fbTrigNewLot   : R_TRIG;                // 新批次上升沿检测实例 / Rising edge detector for the new lot flag
    fbTrigReset    : R_TRIG;                // 复位上升沿检测实例 / Rising edge detector for the reset flag
END_VAR
VAR CONSTANT
    DL_FLOAT_EPS   : REAL := 1.0E-6;        // 浮点判等与判零容差 [无量纲，按比较量量纲同值使用] / Float equality and zero tolerance
    DL_INF_MAX     : REAL := 1.0E30;        // 有限值幅值上限 [无量纲，按各量量纲同值使用] / Finite magnitude upper bound
    DL_LAMBDA_DEF  : REAL := 0.30;          // EWMA 权重默认回退值 [无量纲]，非有限权值时使用 / Default EWMA weight used for non-finite input
    DL_HIST_DEPTH  : INT := 10;             // 历史环缓冲深度 [批]，与结构体数组上界一致 / History ring depth in lots, matching the array bound
    DL_LOT_MAX     : UDINT := 16#FFFF_FFFE; // 批次计数饱和上限 [批]，防累加溢出 / Lot counter saturation limit against overflow
END_VAR

(*------------------------------------------------------------------------------
 * 段 1｜边沿实例无条件周期刷新（红线 R7：严禁置于 IF 或 CASE 分支内）
 *      Unconditional edge refresh, never placed inside IF or CASE branches
 *-----------------------------------------------------------------------------*)
fbTrigNewLot(CLK := bNewLot);
fbTrigReset(CLK := bReset);

(*------------------------------------------------------------------------------
 * 段 2｜瞬时输出与瞬时码预清零（单拍标志在每拍入口清零，出口只置位）
 *      Pre-clear transient outputs and info codes at scan entry
 *-----------------------------------------------------------------------------*)
bCorrected := FALSE;                        // 单拍修正脉冲预清零 [BOOL] / Pre-clear the correction pulse
bAtLimit   := FALSE;                        // 触限标志预清零，本拍按条件重算 [BOOL] / Pre-clear the at-limit flag
uErrInfo   := 0;                            // 瞬时信息码预清零，本拍按条件重算 [码] / Pre-clear the transient info code

(*------------------------------------------------------------------------------
 * 段 3｜参数域修复与 EWMA 权重双向钳位（引脚可在线改，故逐拍重算）
 *      Parameter domain repair and two-sided EWMA weight clamping
 *-----------------------------------------------------------------------------*)
IF fParamMax < fParamMin THEN
    fLimLow  := fParamMax;                  // 域上下对调修复：下限取原上限 [参数单位] / Repaired lower bound takes the original upper
    fLimHigh := fParamMin;                  // 域上下对调修复：上限取原下限 [参数单位] / Repaired upper bound takes the original lower
ELSE
    fLimLow  := fParamMin;                  // 合法下限直通 [参数单位] / Valid lower bound passed through
    fLimHigh := fParamMax;                  // 合法上限直通 [参数单位] / Valid upper bound passed through
END_IF

// 退化域判定：上下限重合时参数被钉死，任何修正都等价于到界，只置 bAtLimit 不另占码位
IF ABS(fLimHigh - fLimLow) <= DL_FLOAT_EPS THEN
    bDomainDeg := TRUE;                     // 参数域无自由度 [BOOL] / Parameter domain has no freedom
    fLimHigh   := fLimLow;                  // 收紧上限与下限对齐，保证 LIMIT 的入参有序 [参数单位] / Tighten the upper bound to keep LIMIT arguments ordered
ELSE
    bDomainDeg := FALSE;                    // 参数域有自由度 [BOOL] / Parameter domain has freedom
END_IF

// EWMA 权重 λ 双向钳位：非有限值回默认、负值钳 0、大于 1 钳 1，均置信息级 1F01
IF (fLambda <> fLambda) OR (ABS(fLambda) > DL_INF_MAX) THEN
    fLambdaEff := DL_LAMBDA_DEF;            // 非有限权值回默认 0.30 [无量纲] / Non-finite weight falls back to the default
    uErrInfo   := 16#0002_1F01;             // 【信息级】λ 越界已钳位 / Info: lambda clamped
ELSIF fLambda < 0.0 THEN
    fLambdaEff := 0.0;                      // 负权值钳到 0，EWMA 冻结在上次值 [无量纲] / Negative weight clamped to zero, EWMA frozen
    uErrInfo   := 16#0002_1F01;             // 【信息级】λ 越界已钳位 / Info: lambda clamped
ELSIF fLambda > 1.0 THEN
    fLambdaEff := 1.0;                      // 大于 1 钳到 1，退化为只看本批 [无量纲] / Weight above one clamped, only this lot used
    uErrInfo   := 16#0002_1F01;             // 【信息级】λ 越界已钳位 / Info: lambda clamped
ELSE
    fLambdaEff := fLambda;                  // 合法权值直通 [无量纲] / Valid weight passed through
END_IF

// 单次修正限幅域修复：取绝对值，非有限值按 0 处理（等效禁止修正，由 1F03 表达）
IF (fCorrectionLim <> fCorrectionLim) OR (ABS(fCorrectionLim) > DL_INF_MAX) THEN
    fCorrLimEff := 0.0;                     // 限幅非有限 → 禁止修正，保守不下发 [参数单位] / Non-finite limit disables correction conservatively
ELSE
    fCorrLimEff := ABS(fCorrectionLim);     // 限幅取绝对值，负号无工程意义 [参数单位] / Absolute limit, sign has no engineering meaning
END_IF

(*------------------------------------------------------------------------------
 * 段 4｜输入有限性体检（NaN 自比较是 IEEE754 唯一可靠的判非数手段）
 *      Input finiteness check, NaN self-comparison is the only reliable test
 *-----------------------------------------------------------------------------*)
bInputsOk := NOT ((fMeasure <> fMeasure) OR (ABS(fMeasure) > DL_INF_MAX)
              OR (fTarget <> fTarget)   OR (ABS(fTarget) > DL_INF_MAX)
              OR (fGainInv <> fGainInv) OR (ABS(fGainInv) > DL_INF_MAX));

(*------------------------------------------------------------------------------
 * 段 5｜首扫装载（R19 唯一合法范式：bInit 初值 FALSE，判据 NOT bInit）
 *      First-scan load, the only accepted pattern for initialisation
 *-----------------------------------------------------------------------------*)
IF NOT bInit THEN
    IF (fParamInit <> fParamInit) OR (ABS(fParamInit) > DL_INF_MAX) THEN
        fParamOut := fLimLow;               // 初始参数非法 → 回退参数域下限 [参数单位] / Non-finite initial parameter falls back to the lower bound
    ELSE
        fParamOut := LIMIT(fLimLow, fParamInit, fLimHigh); // 初始参数钳入参数域 [参数单位] / Initial parameter clamped into the domain
    END_IF
    stHist.fLastParam := fParamOut;         // 历史基准同步，之后一律以历史值为准 [参数单位] / Sync the history baseline used from now on
    stHist.fLastEwma  := 0.0;               // 平滑值清零，bHasEwma 为 FALSE 时不会被使用 [测量单位] / Clear smoothed deviation, unused while the flag is FALSE
    stHist.bHasEwma   := FALSE;             // 首样本标志清零，第一批必走直取路径 [BOOL] / Clear the first-sample flag so the first lot takes over directly
    stHist.nBufIdx    := 0;                 // 环索引归零，第一批写入 1 号槽 [槽] / Ring index reset, the first lot writes slot one
    bInit             := TRUE;              // 首扫完成置位 [BOOL] / First scan completed
END_IF

(*------------------------------------------------------------------------------
 * 段 6｜复位（R19：清 EWMA 与故障，参数保持；复位优先于本拍新故障重锁）
 *      Reset clears EWMA and faults, keeps the parameter, takes priority
 *-----------------------------------------------------------------------------*)
IF fbTrigReset.Q THEN
    uErrFault         := 0;                 // 锁存故障码清零 [码] / Clear the latched fault code
    uErrInfo          := 0;                 // 瞬时信息码清零 [码] / Clear the transient info code
    stHist.bHasEwma   := FALSE;             // 平滑样本作废，下批重新首样本直取 [BOOL] / Invalidate the smoothed sample, next lot takes over directly
    stHist.fLastEwma  := 0.0;               // 平滑值清零 [测量单位] / Clear the smoothed deviation
    stHist.nBufIdx    := 0;                 // 环索引归零，审计从空缓冲重新开始 [槽] / Ring index reset, audit restarts from an empty buffer
    fEwmaDev          := 0.0;               // 平滑偏差出口清零 [测量单位] / Clear the smoothed deviation output
    eState            := E_DL_R2rState.eIdle; // 回空闲态 [枚举] / Back to idle
END_IF

(*------------------------------------------------------------------------------
 * 段 7｜使能撤除：回空闲并保持参数（故障锁存优先于使能撤除，防掩盖故障）
 *      Enable removal returns to idle and holds the parameter, faults win
 *-----------------------------------------------------------------------------*)
IF (NOT bEnable) AND (eState <> E_DL_R2rState.eFault) THEN
    eState := E_DL_R2rState.eIdle;          // 强制回空闲，参数由段 9 派生保持 [枚举] / Force idle, the parameter is held by the mapping section
END_IF

(*------------------------------------------------------------------------------
 * 段 8｜主状态机（红线 R6：ENUM + CASE + ELSE 兜底，五态各有标签）
 *      Main state machine with mandatory ELSE fallback and five labelled states
 *-----------------------------------------------------------------------------*)
CASE eState OF

    E_DL_R2rState.eIdle:                    // 空闲：等使能，不做任何参数动作
        IF bEnable THEN
            eState := E_DL_R2rState.eReady; // 使能到位即进就绪 [枚举] / Enable asserted moves to ready
        END_IF

    E_DL_R2rState.eReady:                   // 就绪：等新批次沿；期间持续体检输入有限性
        IF NOT bInputsOk THEN
            uErrFault := 16#0002_1F10;      // 【故障级】输入非有限值，锁存待复位 / Fault: non-finite input latched until reset
            eState    := E_DL_R2rState.eFault;
        ELSIF fbTrigNewLot.Q THEN
            eState := E_DL_R2rState.eCompute; // 批次沿开启事务 [枚举] / Lot edge opens the transaction
        END_IF

    E_DL_R2rState.eCompute:                 // 计算：偏差 → EWMA → 修正量，本拍算完即转
        IF NOT bInputsOk THEN
            uErrFault := 16#0002_1F10;      // 【故障级】输入非有限值，锁存待复位 / Fault: non-finite input latched until reset
            eState    := E_DL_R2rState.eFault;
        ELSE
            fDev := fMeasure - fTarget;     // 本批原始偏差 [测量单位] / Raw deviation of this lot
            IF NOT stHist.bHasEwma THEN
                fEwmaDev        := fDev;    // 首样本直取，绝不与 0 平均 [测量单位] / First sample taken over directly, never averaged with zero
                stHist.bHasEwma := TRUE;    // 置样本有效标志，后续批次走递推 [BOOL] / Mark the sample valid for subsequent recursion
                uErrInfo        := 16#0002_1F02; // 【信息级】无历史样本，首样本直取 / Info: no history, first sample taken over
            ELSE
                fEwmaDev := fLambdaEff * fDev + (1.0 - fLambdaEff) * stHist.fLastEwma; // EWMA 递推 [测量单位] / EWMA recursion
            END_IF
            stHist.fLastEwma := fEwmaDev;   // 平滑值存档供下批递推 [测量单位] / Archive the smoothed value for the next lot
            fCorr := -fEwmaDev * fGainInv;  // 修正量＝负偏差乘增益倒数 [参数单位] / Correction equals negative deviation times inverse gain
            IF ABS(fCorr) > fCorrLimEff THEN
                fCorr     := LIMIT(-fCorrLimEff, fCorr, fCorrLimEff); // 单次限幅，双向钳位 [参数单位] / Per-lot two-sided clamp
                bAtLimit  := TRUE;          // 修正量触限 [BOOL] / Correction at its limit
                uErrInfo  := 16#0002_1F03;  // 【信息级】修正量达限幅 / Info: correction at the per-lot limit
            END_IF
            eState := E_DL_R2rState.eApply; // 算完立即转回写态，两态各驻留一拍 [枚举] / Move to apply, each state stays exactly one scan
        END_IF

    E_DL_R2rState.eApply:                   // 回写：参数钳入参数域 → 记审计 → 出单拍
        fParamNew := LIMIT(fLimLow, stHist.fLastParam + fCorr, fLimHigh); // 参数域第二重约束 [参数单位] / Domain clamping as the second constraint
        IF (ABS(fParamNew - fLimHigh) <= DL_FLOAT_EPS) OR (ABS(fParamNew - fLimLow) <= DL_FLOAT_EPS) THEN
            bAtLimit := TRUE;               // 参数顶到域边界，只置触限标志不另占码位 [BOOL] / Parameter pinned at a bound, flag only
        END_IF
        IF bDomainDeg THEN
            bAtLimit := TRUE;               // 退化域下任何修正都等价于到界 [BOOL] / Degenerate domain makes every correction a limit hit
        END_IF
        stHist.fLastParam := fParamNew;     // 历史参数推进，出口由段 9 派生 [参数单位] / Advance the historical parameter, mapped in the final section
        stHist.nBufIdx    := stHist.nBufIdx + 1; // 环写指针前进一格 [槽] / Advance the ring write index
        IF stHist.nBufIdx < 1 THEN
            stHist.nBufIdx := 1;            // 下界校验：索引不得小于 1 [槽] / Lower bound guard, index never below one
        ELSIF stHist.nBufIdx > DL_HIST_DEPTH THEN
            stHist.nBufIdx := 1;            // 上界校验：越界即环绕回首槽 [槽] / Upper bound guard, wrap to the first slot
        END_IF
        IF (stHist.nBufIdx >= 1) AND (stHist.nBufIdx <= DL_HIST_DEPTH) THEN
            stHist.afDevBuf[stHist.nBufIdx] := fDev; // 偏差写入环缓冲 [测量单位] / Write the deviation into the ring buffer
        END_IF
        IF uLotCount < DL_LOT_MAX THEN
            uLotCount := uLotCount + 1;     // 批次计数饱和累加，封顶不溢出 [批] / Saturating lot counter
        END_IF
        bCorrected := TRUE;                 // 单拍修正脉冲，下一拍入口由段 2 清零 [BOOL] / Single-scan correction pulse, cleared at the next scan entry
        eState     := E_DL_R2rState.eReady; // 本批事务结束，回就绪等下一批 [枚举] / Transaction finished, back to ready

    E_DL_R2rState.eFault:                   // 故障锁存：参数保持，仅复位沿退出
        bCorrected := FALSE;                // 故障态不再输出修正脉冲 [BOOL] / No correction pulse while faulted
        bAtLimit   := FALSE;                // 故障态触限标志无意义，保持清零 [BOOL] / At-limit flag cleared while faulted

    ELSE                                    // 非法状态兜底：一律回故障态并复用本块最高优先故障码
        uErrFault := 16#0002_1F10;          // 【故障级】非法状态兜底，复用 1F10 / Fault: illegal state fallback reusing 1F10
        eState    := E_DL_R2rState.eFault;  // 强制进故障锁存 [枚举] / Force the latched fault state

END_CASE

(*------------------------------------------------------------------------------
 * 段 9｜出口映射（派生式：信息级码只进 uErrorId，bError 只反映 eFault 态）
 *      Output mapping, info codes never raise the fault flag
 *-----------------------------------------------------------------------------*)
fParamOut := stHist.fLastParam;             // 下发参数恒等于历史生效参数 [参数单位] / Output parameter always mirrors the historical effective value
bError    := (eState = E_DL_R2rState.eFault); // 故障标志只由 eFault 态派生 [BOOL] / Fault flag derived from the fault state only
IF eState = E_DL_R2rState.eFault THEN
    uErrorId := uErrFault;                  // 故障态上报锁存码，不被本拍信息码覆盖 [码] / Report the latched code while faulted
ELSE
    uErrorId := uErrInfo;                   // 运行态上报本拍瞬时信息码 [码] / Report the transient info code while running
END_IF

END_FUNCTION_BLOCK
